(* IEC 61131-3 sources: plcassist-cli/packages/volt-lsp-iec/test-corpus/pro2193/Device/Plc Logic/Application/09 Misc/Library Manager/L_TT1P_TechnologyModules (part 4) *)

(* ---- L_MB1P_TPCALCDIFF.fb ---- *)
FUNCTION_BLOCK L_MB1P_TPCALCDIFF
VAR_INPUT
	XENABLE : BOOL;
	XTPRECEIVED : BOOL;
	LRACTTPPOSIN : LREAL;
	LRSETTPPOSIN : LREAL;
	LRSETMARKDISTANCE : LREAL;
END_VAR
VAR_OUTPUT
	XINITDONE : BOOL;
	XTPRECEIVEDOUT : BOOL;
	LRTPDIFFERENCE : LREAL;
	LRTPDIFFTOTAL : LREAL;
END_VAR
VAR
	XTPRECEIVEDOLD : BOOL;
END_VAR
END_FUNCTION_BLOCK

(* ---- L_MB1P_TPCONVERTTP.fb ---- *)
FUNCTION_BLOCK L_MB1P_TPCONVERTTP
VAR_INPUT
	XENABLE : BOOL;
	XTPRECEIVE : BOOL;
	LRACTTPPOSIN : LREAL;
	LRDELAYACTSET : LREAL;
	LRCYCPOSTPAXIS : LREAL;
	LRCYCPOSTARGETAXIS : LREAL;
	LRCYCLELENGTHTPAXIS : LREAL;
	LRCYCLELENGTHTARGETAXIS : LREAL;
END_VAR
VAR_OUTPUT
	XTPRECEIVED : BOOL;
	LRTPACTPOS : LREAL;
	XERROR : BOOL;
	EERRORID : L_IE1P_Error;
END_VAR
VAR
	LRPOSFIFOX : ARRAY [1..20] OF LREAL := [10(0)];
	LRPOSFIFOREG : ARRAY [1..20] OF LREAL := [10(0)];
	BYCOUNTER : INT := 1;
	LRSTACKDIFFERENCE : LREAL;
	LRTPDELTAINMS : LREAL;
	LRDELTAPCT : LREAL;
	XTPRECEIVEDOLD : BOOL;
	LRPOSDIFFTPAXIS : LREAL;
	IDIRECTION : INT;
	LRACTTPPOSIN_OLD : LREAL;
	XWAIT : BOOL;
	XWAIT_OLD : BOOL;
	LRACTTPPOSIN_INT : LREAL;
	R_TRIG1 : R_TRIG;
	BYCOMPENSATIONCYCLES : BYTE;
	LRDELAYACTSETRESIDUAL : LREAL;
	LRDELTATARGETAXIS : LREAL;
END_VAR
END_FUNCTION_BLOCK

METHOD SEARCHINSTACKNEGATIVE
END_METHOD

METHOD SEARCHINSTACKPOSITIVE
END_METHOD

(* ---- L_MB1P_TPLIMITDIFF.fb ---- *)
FUNCTION_BLOCK L_MB1P_TPLIMITDIFF
VAR_INPUT
	XTPRECEIVED : BOOL;
	LRSETTPDIFFERENCE : LREAL;
	LRSETLIMITMIN : LREAL := -100;
	LRSETLIMITMAX : LREAL := 100;
	LRSETTPWINDOW : LREAL := 2;
END_VAR
VAR_OUTPUT
	XTPRECEIVEDOUT : BOOL;
	XLIMITACTIVE : BOOL;
	XTPINWINDOW : BOOL;
	LRTPDIFFERENCELIM : LREAL;
END_VAR
VAR
	XTPRECEIVEDOLD : BOOL;
	XINITDONE : BOOL;
END_VAR
END_FUNCTION_BLOCK

(* ---- L_MB1P_TPVIRTUALACTPOS.fb ---- *)
FUNCTION_BLOCK L_MB1P_TPVIRTUALACTPOS
VAR_INPUT
	XTPWINDOWOPEN : BOOL;
	XTPRECEIVEDIN : BOOL;
	XMAXTPNOTDETECTED : BOOL;
	LRSETTPPOSIN : LREAL;
	LRACTTPPOSIN : LREAL;
END_VAR
VAR_OUTPUT
	XTPRECEIVEDOUT : BOOL;
	LRACTTPPOS : LREAL;
END_VAR
VAR
	XTPRECEIVEDINOLD : BOOL;
	XFLAGWINDOWOPENANDNOTP : BOOL := FALSE;
	XWINDOWOPENOLD : BOOL;
	XVIRTUALTPACTIVE : BOOL;
END_VAR
END_FUNCTION_BLOCK

(* ---- L_MB1P_WINDERIDENTDIAMETER.fb ---- *)
FUNCTION_BLOCK L_MB1P_WINDERIDENTDIAMETER
VAR_INPUT
	XEXECUTE : BOOL;
	XABORT : BOOL;
	XDANCERMINPOS : BOOL;
	LRACTREELSPEEDIN : LREAL;
	LRACTDANCERPOSIN : LREAL;
	XLINEVELDIAMCALC : BOOL;
	LRSETLINEVELDIAMCALC : LREAL;
	LRMAXDANCERPOS : LREAL;
	LRDANCERMATERIALLENGTH : LREAL;
	LRMAXDIAM : LREAL;
	LRDIAMCALCDIST : LREAL;
	WIDENTDIAMCALCCYCLES : WORD := 1;
	LRTASKCYCLE : LREAL := 0.001;
	LRIDENTVEL : LREAL;
	LRIDENTACC : LREAL;
	LRIDENTDEC : LREAL;
	LRIDENTJERK : LREAL;
END_VAR
VAR_OUTPUT
	XERROR : BOOL;
	EERRORID : WORD;
	XBUSY : BOOL;
	XDONE : BOOL;
	XCOMMANDABORTED : BOOL;
	LRSETREELSPEEDOUT : LREAL;
	LRIDETDIAM : LREAL;
END_VAR
VAR
	WSTATE : WORD;
	LRTASKCYCLE_INT : LREAL := 0.001;
	LRMAXDIAM_INT : LREAL;
	LRREELSPEEDFAKTOR_INT : LREAL;
	LRMAXDANCERPOS_INT : LREAL;
	LRDANCERMATERIALLENGTH_INT : LREAL;
	XLINEVELDIAMCALC_INT : BOOL;
	LRREELSPEEDOUT_INT : LREAL;
	LRACTREELDIST_INT : LREAL;
	LRACTDIST_INT : LREAL;
	LRPROFGENDIST_INT : LREAL;
	LRSETDIST_INT : LREAL;
	LRSETDISTCALCDIAM_INT : LREAL;
	LRPROFGENSTARTPOSIDENTDIAM_INT : LREAL;
	LRPROFGENENDPOSIDENTDIAM_INT : LREAL;
	LRRAMPGENDECDIST : LREAL;
	XRAMPGENHALT : BOOL;
	XIDENTSTARTVALUESVALID : BOOL;
	XIDENTENDVALUESVALID : BOOL;
	LRDANCERPOSSTARTIDENT : LREAL;
	LRDANCERPOSENDIDENT : LREAL;
	LRLINEVELSTARTIDENT : LREAL;
	LRLINEVELENDIDENT : LREAL;
	LRLINEDIST : LREAL;
	LRWNDPOSSTARTIDENT : LREAL;
	LRWNDPOSENDIDENT : LREAL;
	LRIDETNWINDDIST : LREAL;
	XERROR_INVALIDMAXDIAM : BOOL;
	XERROR_INVALIDDANCERMATERIALLENGTH : BOOL;
	XERROR_ACTDANPOSBIGGERMAXDANPOS : BOOL;
	XERROR_ACTDANPOSBIGGERMAXDANPOS_TMP : BOOL;
	XEXECUTE_OLD : BOOL;
	XABORT_OLD : BOOL;
	FB_RAMPGENERATOR1 : L_MC1P_RampGenerator;
END_VAR
END_FUNCTION_BLOCK

METHOD CALL_ERRORHANDLER
END_METHOD

METHOD CALL_FBMETHODS
END_METHOD

METHOD CALL_FB_RAMPGENERATOR
END_METHOD

METHOD CALL_OUTPUT
END_METHOD

METHOD CALL_RESETCOMMANDS
END_METHOD

METHOD CALL_RESETOUTPUT
END_METHOD

METHOD CALL_STATEMACHINE
END_METHOD

(* ---- L_MB1P_WINDERSYNCHRONISELINE.fb ---- *)
FUNCTION_BLOCK L_MB1P_WINDERSYNCHRONISELINE
VAR_INPUT
	XENABLE : BOOL;
	XSYNCLINEVEL : BOOL;
	XLOADSTARTREELSPEED : BOOL;
	LRSTARTREELSPEED : LREAL;
	LRGROUNDREELSPEED : LREAL;
	LRCYCLINEVEL : LREAL := 0;
	LRSETDIAMETER : LREAL;
	LRACC : LREAL := 1000;
	LRDEC : LREAL := 1000;
	LRJERK : LREAL := 100000;
	XMATERIALFEEDING : BOOL := FALSE;
END_VAR
VAR_OUTPUT
	XERROR : BOOL;
	EERRORID : WORD;
	XBUSY : BOOL;
	XSYNCHRONISED : BOOL;
	XACCDECSYNC : BOOL;
	LRSETREELSPEEDOUT : LREAL;
END_VAR
VAR
	WSTATE : WORD;
	LRREELSPEEDOUT_INT : LREAL;
	FB_RAMPGENERATOR1 : L_MC1P_RampGenerator;
	XENABLE_OLD : BOOL;
	XMATERIALFEEDING_OLD : BOOL;
	LRSCALEFAKTOR : LREAL;
	LRSCALEFAKTORABS : LREAL;
	WPARMODE : WORD;
	XTMP : BOOL;
END_VAR
END_FUNCTION_BLOCK

METHOD CALL_ERRORHANDLER
END_METHOD

METHOD CALL_FBMETHODS
END_METHOD

METHOD CALL_FB_RAMPGENERATOR
END_METHOD

METHOD CALL_OUTPUT
END_METHOD

METHOD CALL_RESETCOMMANDS
END_METHOD

METHOD CALL_RESETOUTPUT
END_METHOD

METHOD CALL_SETPARMODE
END_METHOD

METHOD CALL_STATEMACHINE
END_METHOD

(* ---- L_T01S_PHASECORRECTIONVEL.fb ---- *)
FUNCTION_BLOCK L_T01S_PHASECORRECTIONVEL
VAR_INPUT
	XENABLE : BOOL;
	XEXECUTECORRECTION : BOOL;
	LRCYCSETVEL : LREAL;
	LRSETCORRECTION : LREAL;
	LRCORRECTIONDISTANCE : LREAL;
END_VAR
VAR_OUTPUT
	XBUSY : BOOL;
	XCORRECTIONBUSY : BOOL;
	LRSETVELOUT : LREAL;
	LRSETCORRVELOUT : LREAL;
	LRSETPOSCORROUT : LREAL;
	XERROR : BOOL;
	EERRORID : L_IE1P_Error;
END_VAR
VAR
	LRDELTAPOSTOTAL : LREAL;
	LRMASTERDISTANCE : LREAL;
	LRPOSITIONSET : LREAL;
	LRPOSITIONNORMED : LREAL;
	LRPOSITIONOUTNORMED : LREAL;
	LRDELTAPOSCORRECTION : LREAL;
	LRPOSITIONSETOLD : LREAL;
	BYSTEPPER : BYTE;
	LRCORRECTIONDISTANCELOCAL : LREAL;
	LRCORRECTIONLOCAL : LREAL;
	LRDELTAPOSOUT : LREAL;
	XEXECUTECORRECTIONINTERN : BOOL;
	LRTASKCYCLE : LREAL;
	XINIT : BOOL := TRUE;
	INTEGRATE1 : L_USPP_Integrate;
END_VAR
END_FUNCTION_BLOCK

(* ---- L_TF1P_ADDPROFILEPICKANDPLACE.fb ---- *)
FUNCTION_BLOCK L_TF1P_ADDPROFILEPICKANDPLACE
VAR_INPUT
	XENABLE : BOOL;
	XEXECUTEPICKANDPLACE : BOOL;
	XADDPROFILE : BOOL;
	XRESETTARGETSTACK : BOOL;
	XACKPATHHALT : BOOL;
	XABORT : BOOL;
	XNOTCOORDINATEDSTOPALL : BOOL;
	XSINGLESTEP : BOOL;
	LRGRIPPERTIME : LREAL;
	LRPATHJERK : LREAL;
	LRNUMTASKCYCLESBEFOREEXECUTENEXTPROFILE : LREAL := 50;
	XCALCPROFILEMOVEPATH : BOOL;
END_VAR
VAR_OUTPUT
	XERROR : BOOL;
	XWARNING : BOOL;
	EERRORID : L_IE1P_Error;
	XBUSY : BOOL;
	XACTIVE : BOOL;
	XDONE : BOOL;
	XCOMMANDABORTED : BOOL;
	XENDOFPROFILE : BOOL;
	XTARGETSTACKISFULL : BOOL;
	XPATHHOLD : BOOL;
	XPROFILEINPREPARATION : BOOL;
	ISETPROFILENOOUT : INT;
	IPROFILEPOINTPASSED : INT;
	ITARGETPROFILEPOINT : INT;
	ALRTARGETPOSITION : ARRAY [1..12] OF LREAL;
	ESETSEGMENTTYPEOUT : L_MC4P_SegmentType;
	BYNUMOFPOINTSINPROFILE : BYTE;
	BYNUMOFHALTINPROFILE : BYTE;
	LRPATHPREPARATIONTIME : LREAL;
	LRPRECALCPROFILETIME : LREAL;
	XPROFILERESTTIMEVALID : BOOL;
	LRPROFILERESTTIME : LREAL;
	LRINTERRUPTPATHACC : LREAL;
	XLASTACTIVESEGMENT : BOOL;
	XNOACTIVESEGMENT : BOOL;
	XGRIPPERCTRLACTIVE : BOOL;
	XPULSEGRIPPER : BOOL;
	XPATHINTERRUPTOUT : BOOL;
	PAFB_MOVELINABS : POINTER TO ARRAY [1..10] OF L_MC4P_MoveLinearAbsolute_Internal;
	IMOVEPPNO : INT;
	IMOVELINNO : INT;
	PAFB_MOVELINABS1 : POINTER TO ARRAY [1..10] OF L_MC4P_MoveLinearAbsolute_Internal;
	PAFB_MOVELINABS2 : POINTER TO ARRAY [1..10] OF L_MC4P_MoveLinearAbsolute_Internal;
	PAFB_MOVELINABS3 : POINTER TO ARRAY [1..10] OF L_MC4P_MoveLinearAbsolute_Internal;
	XWAITDISABLEMOVECONTPATH : BOOL;
END_VAR
VAR_IN_OUT
	FB_EXTERNALMEMORY : L_MC4P_PickAndPlaceMemory;
	AXESGROUP : AXES_GROUP_KIN;
	ASCPROFILEPAR : ARRAY [1..10] OF L_TT1P_scProfilePar;
END_VAR
VAR
	LWTCHECKSUM_INT : LWORD;
	WSTATE : WORD;
	XSTATEMASHINEBUSY : BOOL;
	XSTATEMASHINEWAIT : BOOL;
	XSTATEMASHINEPATHHOLD : BOOL;
	XMOVEPAPSTATUSSEPPERENTRY : BOOL;
	WMOVEPAPSTATUSSEPPER_OLD : WORD;
	WMOVEPAPSTATUSSEPPER : WORD;
	REQUESTSINFO : DWORD;
	REQUESTSINFO_OLD : DWORD;
	DWRTRIG : DWORD;
	DWFTRIG : DWORD;
	EBUFFERMODEBLENDING_INT : MC_BUFFER_MODE := MC_BUFFER_MODE.mcBlendingLow;
	LRTEMP1 : LREAL;
	LRTEMP2 : LREAL;
	IDX1 : INT;
	IDX2 : INT;
	IDX3 : INT;
	UIDX1 : UINT;
	WDX1 : WORD;
	TTMP1 : TIME;
	WTMP1 : WORD;
	IFOR : INT;
	IFOREND : INT;
	ALRTARGETPOSTMP : ARRAY [1..12] OF LREAL;
	XCOUNTUPPROFILENOOUT : BOOL;
	XERRORINVALIDPROFILE : BOOL;
	XERROR_INVALIDCOORDSYSTEM : BOOL;
	XERROR_INVALIDTARGET : BOOL;
	XERROR_INVALIDPATHPAR : BOOL;
	XWARNING_TARGETSTATCKISFULL : BOOL;
	XWARNING_NOTREADYFORADDPROFILE : BOOL;
	XERROR_FB_MOVEPICKANDPLACE : BOOL;
	EERRORID_FB_MOVEPICKANDPLACE : L_IE1P_Error;
	XERROR_INTERNAL : BOOL;
	XERRORINTERNAL_INVALIDPPFBACTIVE : BOOL;
	WINTERNALERRORID_INT : WORD;
	XSINGLESTEP_LOCK : BOOL;
	LRGRIPPERTIME_LOCK : LREAL;
	XCALLFM : BOOL;
	LRTASKCYCLE : LREAL;
	LRTASKCYCLE_INV : LREAL;
	LRTIMEBEFOREEXECUTENEXTPROFILE : LREAL;
	FB_STACKTARGET : L_MC1P_StackControlArray := STRUCT(iMaxLegth := ciNumOfTargetInArray);
	ALRTARGETGRIPPERTIME : ARRAY [1..ciNumOfTargetInArray] OF LREAL;
	ALRPATHJERK : ARRAY [1..ciNumOfTargetInArray] OF LREAL;
	AXTARGETGRIPPERTIMEVALID : ARRAY [1..ciNumOfTargetInArray] OF BOOL;
	AXSINGLESTEP_INT : ARRAY [1..ciNumOfTargetInArray] OF BOOL;
	XNEWTARGET : BOOL;
	XAXESGROUPNOTREADYFORMOTION : BOOL;
	XNEXTPROFILEVALID : BOOL;
	XMOVEPPPATHINTERRUPTOUT : BOOL;
	IGRIPPERMOVEPPNO : INT;
	XPREPARENEXTPROFILE : BOOL;
	XPATHACTIVE_INT : BOOL;
	XPATHBUSY_INT : BOOL;
	XPATHDONE_INT : BOOL;
	XPATHHOLD_INT : BOOL;
	XPATHHOLDONENDHALT_INT : BOOL;
	XPATHINTERRUPTOUT_INT : BOOL;
	XPATHCOMMANDABORTED_INT : BOOL;
	XCOMMANDABORTED_INT : BOOL;
	XCOMMANDABORTE_INT : BOOL;
	XPROFILEINPREPARATION_INT : BOOL;
	LRPRECALCRESTTIMEALLSEGMENTS_INT : LREAL;
	XPRECALCPROFILERESTTIMEALLSEGMENTSVALID_INT : BOOL;
	XPRECALCPROFILERESTTIMEVALID_INT : BOOL;
	LRPRECALCPROFILERESTTIME_INT : LREAL;
	LRIPOTIME : LREAL;
	LRPATHPREPARATIONTIME_INT : LREAL;
	INUMOFACTIVEPATHSEGMENT_INT : INT;
	ICNTRACKPATHHALT_INT : INT;
	XVALIDSTARTPOS : BOOL;
	XSTARTPOINTINHALT_INT : BOOL;
	ALRSTARTPOS_INT : ARRAY [1..12] OF LREAL;
	ESTARTCOORDSYSTEM_INT : L_MC4P_CoordSystem;
	LRSTARTBLENDINGRADIUS_INT : LREAL;
	XSAVEPROFILE_INT : BOOL;
	ISAVEPROFILEEXECUTED_INT : INT;
	ISAVEPROFILESTACKSTARTPOS_INT : INT;
	ISAVEPROFILESTACKLEGTH_INT : INT;
	FB_STACKMOVEPICKANDPALCE : L_MC1P_StackControlArray := STRUCT(iMaxLegth := ciNumOfFBMovePickAndPlace);
	AIPROFILENOSTATIC : ARRAY [1..ciNumOfFBMovePickAndPlace] OF INT;
	FB_MOVEPICKANDPLACE : ARRAY [1..ciNumOfFBMovePickAndPlace] OF L_MB1P_MovePickAndPlaceState;
	CINUMOFTARGETINARRAY : INT := 10;
	CINUMOFTARGETINARRAYSETWARNING : INT := 8;
	CINUMOFFBMOVEPICKANDPLACE : INT := 3;
	EBUFFERMODEBLENDING : MC_BUFFER_MODE;
	LWTCHECKSUM : LWORD;
END_VAR
END_FUNCTION_BLOCK

METHOD CALL_ALLOCPOINTADR
END_METHOD

METHOD CALL_CALCPROFILETIME
END_METHOD

METHOD CALL_DISABLEMOVECONTPATH
VAR_IN_OUT
	AXESGROUP : AXES_GROUP_KIN;
END_VAR
END_METHOD

METHOD CALL_ERRORHANDLER
END_METHOD

METHOD CALL_FBMETHODS
END_METHOD

METHOD CALL_FB_MOVEPICKANDPLACE
END_METHOD

METHOD CALL_FB_MOVEPICKANDPLACE_STATUS
END_METHOD

METHOD CALL_GRIPPERCONTROL
END_METHOD

METHOD CALL_OUTPUT
END_METHOD

METHOD CALL_REQUESTS_EXT
END_METHOD

METHOD CALL_RESETCOMMANDS
END_METHOD

METHOD CALL_RESETOUTPUT
END_METHOD

METHOD CALL_STATEMACHINE
END_METHOD

METHOD CALL_ABORTPROFILE
END_METHOD

METHOD CALL_READSTARTPOSITION
END_METHOD

METHOD CALL_SAVEPROFILE
END_METHOD

METHOD CALL_TARGETSTAICPOSSTACK
END_METHOD

METHOD CALL_SETPROFILE
END_METHOD

METHOD GET_ALRINTERMEDIANTEPOINT
VAR_IN_OUT
	ALRINTERMEDIANTEPOINT : ARRAY [1..12] OF LREAL;
END_VAR
END_METHOD

METHOD CALL_INIT
END_METHOD

METHOD CALL_S000_CYCLIC
END_METHOD

(* ---- L_TF1P_REGISTERCONTROLBASE.fb ---- *)
FUNCTION_BLOCK L_TF1P_REGISTERCONTROLBASE
VAR_INPUT
	XENABLE : BOOL;
	XSYNCPOS : BOOL;
	LRVELIN : LREAL;
	LRACTSETPOSSLAVE : LREAL;
	XMARKRECEIVE : BOOL;
	ETPMODE : L_TF1P_TpMode;
	LRCYCPOSEXTENCODER : LREAL;
	LRCYCLELENGTHEXTENCODER : LREAL;
	LRACTMARKPOSIN : LREAL;
	XLOADREGPOS : BOOL;
	LRLOADREGPOS : LREAL;
	LRMARKSENSORPOS : LREAL;
	LRMARKDIST : LREAL;
	LRMAXCORRNEG : LREAL;
	LRMAXCORRPOS : LREAL;
	ESOURCEFORCORRWINDOW : L_TT1P_SourceForCorrWindow;
	LRUPPERCORRPOS : LREAL;
	LRLOWERCORRPOS : LREAL;
	DNNUMAXISY : DWORD;
	DNDENAXISY : DWORD;
	XSYNCHRONISED : BOOL;
	LRTPAXISCOMPFACTOR : LREAL;
	LRTPAXISDELAYCYCLE : LREAL;
END_VAR
VAR_OUTPUT
	LRPOSOUT : LREAL;
	LRACTVEL : LREAL;
	XERROR : BOOL;
	WERRORID : WORD;
	XLIMITACTIVE : BOOL;
	LRACTMARKERROR : LREAL;
	LRACTMARKDIST : LREAL;
	XINITDONE : BOOL;
	XCORRACTIVE : BOOL;
	XMARKRECEIVED : BOOL;
	LRREGMARKPOS : LREAL;
	XCORRNEXTCYCLE : BOOL;
END_VAR
VAR_IN_OUT
	MASTERAXIS : AXIS_REF;
	SLAVEAXIS : AXIS_REF;
END_VAR
VAR
	SPEEDTOPOSINTEGRATE : L_MC1P_IntegrateAxis;
	TPLIMITDIFF : L_MB1P_TpLimitDiff;
	FB_ADDOFFSET : L_MC1P_AddOffsetCyclic;
	TPCALCDIFF : L_MC1P_TpCalcDiff;
	CONVERTTPPOSITION : L_TT1P_CalculateTPOnMaterialPos := STRUCT(xNoMarkStack := TRUE);
	DISTCORRECTIONWINDOW : L_MB1P_DistCorrectionWindow;
	LRGEARINGFAKTOR : LREAL := 1.0;
	XERROR_TM : BOOL;
	EERRORID_TM : L_IE1P_Error;
	LRTPDIFFERENCE_INT : LREAL;
	XLOADMARKSENSORPOS_OLD : BOOL;
	XTPRECEIVED_OLD : BOOL;
	LRMARKWINDOWSIZE_INT : LREAL;
	XTPINWINDOW : BOOL;
	LRPOS_INT : LREAL;
	XTPRECEIVEDOUT_INT : BOOL;
	LRTPACTPOSITION_INT : LREAL;
	LRTPDIFFERENCELIM_INT : LREAL;
	LROFFSETPOSCTRL_INT : LREAL;
	LRPOSOUT_INT : LREAL;
	LRVELOUT_INT : LREAL;
	XCORRACTIVE_INT : BOOL;
	XINIT : BOOL := TRUE;
	XTPCORRECTIONACTIVE : BOOL := FALSE;
	LRTPAXISSETPOS : LREAL;
	LRMARKDIST_INT : LREAL;
	XZERO : BOOL;
	XHOMINGDONE : BOOL;
	XSTARTREFERENCEACTIVE : BOOL;
	XHOMINGACTIVE : BOOL := FALSE;
	XMARKDISTCHANGED : BOOL;
	XENABLE_OLD : BOOL;
	XTPRECEIVEDOUT_INTOLD : BOOL;
	XSTARTFIRSTCORRECTION : BOOL;
	LRTPDIFFERENCELIM2_INT : LREAL;
	XCORRECTIONBUSYOLD : BOOL;
	LRTPACTPOSIN_OLD : LREAL;
	LRTPSETPOSIN_OLD : LREAL;
	LRCYCLELENGTH : LREAL;
	ICOUNTER : INT := 0;
	LRSETPOSITIONOLD : LREAL;
	LRCYCLELENGTHTP : LREAL;
	LRTPACTPOSITIONOLD : LREAL;
	L_MB1P_CHECKMODULOOVERRUNSETPOS : L_MB1P_CheckModuloOverrun;
	L_MB1P_CHECKMODULOOVERRUNACTPOS : L_MB1P_CheckModuloOverrun;
	BYCYCLECOUNT_INT : BYTE;
	BYCYCLECOUNTREG_INT : BYTE;
	BYSTATE : BYTE;
	ABYCYCLECOUNT : ARRAY [0..5] OF BYTE;
	BYCYCLECOUNTSUM : BYTE;
	XFIRSTTOUCHPROBE : BOOL := TRUE;
	XCORRBASEDONMASTERPOS_INT : BOOL := FALSE;
	XTPCALCDIFFTPRECEIVEDOLD : BOOL;
	LRTPDIFFERENCECOMP_INT : LREAL;
	LRTPAXISACTPOS : LREAL;
	LRTPAXISACTVELOCITY : LREAL;
	LRTPAXISCYCLELENGTH : LREAL;
	LRCYCREGISTERPOSINT : LREAL;
	LRTPACTPOSITION_ORIGINAL : LREAL;
	LRREGISTERTOUCHPROBEDIFFERENCE : LREAL;
	LRAXISTOUCHPROBEDIFFERENCE : LREAL;
END_VAR
END_FUNCTION_BLOCK

METHOD CALL_CALCACTMARKDIST
END_METHOD

METHOD CALL_CORRECTIONPOS
END_METHOD

METHOD CALL_ENABLEREGISTERCONTROL
END_METHOD

METHOD CALL_ERRORHANDLER
END_METHOD

METHOD CALL_FB
END_METHOD

METHOD CALL_GEARING
END_METHOD

METHOD CALL_INPUT
END_METHOD

METHOD CALL_LIMIT
END_METHOD

METHOD CALL_MARKDISTCHANGE
END_METHOD

METHOD CALL_NOTENABLE
END_METHOD

METHOD CALL_OUTPUT
END_METHOD

METHOD CALL_RESET
END_METHOD

METHOD CALL_TOUCHPROBE
END_METHOD

METHOD CALL_TOUCHPROBESOURCE
END_METHOD

METHOD GET_ACTUALMARKDIST : LREAL
END_METHOD

METHOD GET_CORRREGPOS : LREAL
END_METHOD

METHOD GET_INTEGRATORREGPOS : LREAL
END_METHOD

METHOD GET_MARKERRORUNLIMITED : LREAL
END_METHOD

METHOD GET_MARKPOSITIONINREGISTER : LREAL
END_METHOD

METHOD GET_MARKRECEIVEUNLIMITED : BOOL
END_METHOD

METHOD GET_REGISTERINPUTVEL : LREAL
END_METHOD

METHOD GET_SETVELOCITYREGISTER : LREAL
END_METHOD

METHOD SET_CORRECTIONONMASTERPOS
VAR_INPUT
	XCORRBASEDONMASTER : BOOL;
END_VAR
END_METHOD

(* ---- L_TF1P_REGISTERCONTROLSTATE.fb ---- *)
FUNCTION_BLOCK L_TF1P_REGISTERCONTROLSTATE EXTENDS L_TF1P_RegisterControlBase
VAR_INPUT
	LRACTOFFSETMASTERIN : LREAL;
	LRACTOFFSETSLAVEIN : LREAL;
	XTEACHMARKWINDOW : BOOL;
	LRMARKWINDOWSIZE : LREAL;
	LRSETOFFSETMARKWINDOW : LREAL;
	DWMAXNUMBERVIRTUALMARKS : DWORD;
	LRGEARFACTORCORRGAIN : LREAL;
	LRMAXGEARFACTORCORR : LREAL;
	LRSENSORTOOLDISTANCE : LREAL;
	XGEARFACTORCORR : BOOL;
	XGEARFACTORCORRHOLD : BOOL;
	XENABLETOOLCORRECTION : BOOL;
END_VAR
VAR_OUTPUT
	XMARKWINDOWOPEN : BOOL;
	XMARKOUTOFWINDOW : BOOL;
	XMARKNOTDETECTED : BOOL;
	XMARKWINDOWTEACHED : BOOL;
	LRAVERAGEGEARFACTORCORR : LREAL;
	XGEARFACTORCORRLIMITED : BOOL;
END_VAR
VAR
	MARKWINDOW : L_MB1P_MarkWindowRelative;
	MARKSTACK : L_MB1P_MarkStack;
	TPVIRTUALACTPOS : L_MB1P_TpVirtualActPos;
	LRMARKSTACKLENGTH : LREAL;
	LRTPDIFFERENCELIMITOUT_INT : LREAL;
	XTPRECEIVESTACKOUT_INT : BOOL;
	XTPNOTDETECTED_INT : BOOL;
	XMAXTPNOTDETECTED : BOOL;
	LRGEARFACTORINTEGRATOR : LREAL;
	LRGEARFACTORGAIN : LREAL := 1;
	LRGEARFACTORNUMERATORCORR : LREAL;
	LRGEARFACTORNUMERATORCORRLIMITED : LREAL;
	LRGEARFACTORDENOMINATOR : LREAL;
	LRGEARFACTORNUMERATOR : LREAL;
	LCORRECTIONVELIN : LREAL;
	LRDELTAGEARFACTORCORR : LREAL;
	XTPSENSORTEACHEDOLD : BOOL;
	XTPSENSORTEACHEDATLASTMARK : BOOL;
	XCALCMARKDISTINITIALISED : BOOL;
	XTEACHTPSENSOROLD : BOOL;
	LRTPDEADTIMEDIFF : LREAL;
	XTPRECEIVEDOUTOLD_INT : BOOL;
	XMARKSTACKTPRECEIVEDOUTOLD : BOOL;
	LRTPACTPOSITIONREGISTER_INT : LREAL;
	XTPRECEIVEDOUTREGISTER_INT : BOOL;
	XTPRECEIVEDOUTCALCERROR_INT : BOOL;
	LRTPACTPOSMARKWINDOWIN_INT : LREAL;
	LRMASTERACTPOSITIONOLD_INT : LREAL;
END_VAR
END_FUNCTION_BLOCK

METHOD CALL_AVERAGETPDIFF
END_METHOD

METHOD CALL_CALCACTMARKDIST
END_METHOD

METHOD CALL_CORRECTIONPOS
END_METHOD

METHOD CALL_ENABLEREGISTERCONTROL
END_METHOD

METHOD CALL_ERRORHANDLER
END_METHOD

METHOD CALL_FB
END_METHOD

METHOD CALL_INPUT
END_METHOD

METHOD CALL_LIMIT
END_METHOD

METHOD CALL_MARKDISTCHANGE
END_METHOD

METHOD CALL_MARKREGISTER
END_METHOD

METHOD CALL_MARKWINDOW
END_METHOD

METHOD CALL_NOTENABLE
END_METHOD

METHOD CALL_OUTPUT
END_METHOD

METHOD CALL_RESET
END_METHOD

METHOD CALL_TOUCHPROBE
END_METHOD

METHOD CALL_TOUCHPROBESOURCE
END_METHOD

METHOD CALL_VIRTUALACTPOS
END_METHOD

METHOD GET_ACTMARKERRORLIMITED : LREAL
END_METHOD

METHOD GET_MARKRECEIVEDLIMITED : BOOL
END_METHOD

METHOD GET_MARKWINDOWCOMP : BOOL
END_METHOD

METHOD GET_LRMARKSTACKLENGTH : LREAL
END_METHOD

(* ---- L_TF1P_SYNCDRIVEPOSBASE.fb ---- *)
FUNCTION_BLOCK L_TF1P_SYNCDRIVEPOSBASE
VAR_INPUT
	XENABLE : BOOL;
	LRCYCMASTERPOS : LREAL;
	LRCYCMASTERVEL : LREAL;
	LRCYCMASTERACC : LREAL;
	XLOADSTARTSLAVEPOS : BOOL := FALSE;
	LRSTARTSLAVEPOS : LREAL;
	XLOADGEARBOXPOS : BOOL;
	LRLOADGEARBOXPOS : LREAL;
	DWNUMERATOR : DWORD := 1;
	DWDENOMINATOR : DWORD := 1;
	LRSETOFFSET : LREAL;
END_VAR
VAR_OUTPUT
	XERROR : BOOL;
	EERRORID : L_IE1P_Error;
	XBUSY : BOOL;
	LRSETSLAVEPOSOUT : LREAL;
	LRSETSLAVEVELOUT : LREAL;
	LRSETSLAVEACCOUT : LREAL;
	LRSETGEARBOXPOSOUT : LREAL;
	LROFFSET : LREAL;
END_VAR
VAR_IN_OUT
	MASTERAXIS : AXIS_REF;
	SLAVEAXIS : AXIS_REF;
END_VAR
VAR
	LRSCALING_INT : LREAL := 1;
	LRGEARBOXSTARTPOSOUT_INT : LREAL;
	LRSETMASTERVEL_INT : LREAL;
	LRSETMASTERVEL_OLD : LREAL;
	LRSETMASTERACC_INT : LREAL;
	DWDENOMINATOR_INT : DWORD := 1;
	XENABLE_OLD : BOOL;
	WAXESMODE : WORD;
	ESTATE : L_TF1P_States := L_TF1P_States.INIT;
	ESTATE_OLD : L_TF1P_States := L_TF1P_States.INIT;
	XSTATEENTRY : BOOL;
	XENABLEGEARBOX : BOOL;
	FB_ADDOFFSETCYCLIC : L_MC1P_AddOffsetCyclic;
	FB_GEARBOXPOSITION : L_MB1P_GearboxPosition;
	FB_AXISCONVERTER : L_MC2P.L_MC2P_AxisConverterBase;
	LRLOADGEARBOXPOS_INT : LREAL;
	LRSETGEARBOXPOSOUT_INT : LREAL;
	LRSETGEARBOXPOSOUT_OLD : LREAL;
END_VAR
END_FUNCTION_BLOCK

METHOD CALL_AXESMODE
END_METHOD

METHOD CALL_ERRORHANDLER
END_METHOD

METHOD CALL_FBMETHODS
END_METHOD

METHOD CALL_FBMETHODS_FMDISABLE
END_METHOD

METHOD CALL_FB_ADDOFFSETCYCLIC
END_METHOD

METHOD CALL_FB_ADDOFFSETCYCLIC_INPUT
END_METHOD

METHOD CALL_FB_AXISCONVERTER
END_METHOD

METHOD CALL_FB_AXISCONVERTER_INPUT
END_METHOD

METHOD CALL_FB_GEARBOXPOSITION
END_METHOD

METHOD CALL_FB_GEARBOXPOSITION_INPUT
END_METHOD

METHOD CALL_FB_GEARBOXPOSITION_LOADGEARBOXPOS
END_METHOD

METHOD CALL_LOADSLAVESTARTPOS
END_METHOD

METHOD CALL_OUTPUT
END_METHOD

METHOD CALL_OUTPUT_OFFSET
END_METHOD

METHOD CALL_OUTPUT_SETSLAVEOUT
END_METHOD

METHOD CALL_RESETCOMMANDS
END_METHOD

METHOD CALL_RESETFM
END_METHOD

METHOD CALL_RESETOUTPUT
END_METHOD

METHOD CALL_STATEMASHINE
END_METHOD

METHOD CALL_S000_CYCLIC
END_METHOD

METHOD CALL_S001_INIT
END_METHOD

METHOD CALL_S010_READY
END_METHOD

METHOD CALL_S200_SYNCHRON
END_METHOD

METHOD CALL_S998_ERROR
END_METHOD

(* ---- L_TF1P_SYNCDRIVEPOSHIGH.fb ---- *)
FUNCTION_BLOCK L_TF1P_SYNCDRIVEPOSHIGH EXTENDS L_TF1P_SyncDrivePosState
VAR_INPUT
	XSYNCINSTANT : BOOL;
	XSYNCPOSRESTORE : BOOL;
	XLOADOFFSET : BOOL;
	EOFFSETDIRECTION : L_TF1P_Direction;
	EOFFSETPROFILETYPE : L_TF1P_ProfileType := 0;
	LROFFSETVELPOS : LREAL := 100.0;
	LROFFSETVELNEG : LREAL := 100.0;
	LROFFSETACCDEC : LREAL := 1000.0;
	ESYNCDIRECTION : L_TF1P_SyncDirection := L_TF1P_SyncDirection.mcShortestWay;
	ESYNCMODE : L_TF1P_SyncMode := L_TF1P_SyncMode.ramp_dist;
	LRSYNCINTIME : LREAL := 5;
	LRSYNCOUTTIME : LREAL := 5;
	LRSYNCVEL : LREAL := 100;
	LRSYNCACC : LREAL := 1000.0;
	LRSYNCDEC : LREAL := 1000.0;
	LRSYNCJERK : LREAL := 10000000000.0;
	XLOADCLUTCHOFFSET : BOOL := FALSE;
	LRLOADCLUTCHOFFSET : LREAL := 0;
END_VAR
VAR_OUTPUT
	XSETOFFSETBUSY : BOOL;
	XSETOFFSETDONE : BOOL;
	LROFFSETSYNCPOS : LREAL;
END_VAR
VAR
	LRLOADOFFSET_INT : LREAL := 0;
	XSYNCINSTANT_OLD : BOOL;
	FB_SIMPLEPOSSETOFFSETSLAVE : L_MB1P_SimplePosSetOffset;
	FB_SIMPLEPOSSETOFFSETSYNC : L_MB1P_SimplePosSetOffset;
	LRSYNCOFFSET : LREAL;
END_VAR
END_FUNCTION_BLOCK

METHOD CALL_ERRORHANDLER
END_METHOD

METHOD CALL_FBMETHODS
END_METHOD

METHOD CALL_FBMETHODS_FMDISABLE
END_METHOD

METHOD CALL_FB_ADDOFFSETCYCLIC_INPUT
END_METHOD

METHOD CALL_FB_CLUTCHEXTENDEDBASE_INPUT
END_METHOD

METHOD CALL_FB_SIMPLEPOSSETOFFSETSLAVE
END_METHOD

METHOD CALL_FB_SIMPLEPOSSETOFFSETSLAVE_INPUT
END_METHOD

METHOD CALL_FB_SIMPLEPOSSETOFFSETSYNC
END_METHOD

METHOD CALL_FB_SIMPLEPOSSETOFFSETSYNC_INPUT
END_METHOD

METHOD CALL_OUTPUT
END_METHOD

METHOD CALL_OUTPUT_OFFSET
END_METHOD

METHOD CALL_OUTPUT_SIMPLEPOS
END_METHOD

METHOD CALL_RESETCOMMANDS
END_METHOD

METHOD CALL_RESETOUTPUT
END_METHOD

METHOD CALL_SIMPLEPOS_OFFSET
END_METHOD

METHOD CALL_S001_INIT
END_METHOD

(* ---- L_TF1P_SYNCDRIVEPOSSTATE.fb ---- *)
FUNCTION_BLOCK L_TF1P_SYNCDRIVEPOSSTATE EXTENDS L_TF1P_SyncDrivePosBase
VAR_INPUT
	XSYNCPOS : BOOL;
	XSYNCOUTINSTANT : BOOL;
	XTRIMPOS : BOOL;
	XTRIMNEG : BOOL;
	XRESETTRIM : BOOL;
	LRCYCSLAVEPOS : LREAL;
	LRCYCSLAVEVEL : LREAL;
	LRCYCSLAVEACC : LREAL;
	LRTRIMVELPOS : LREAL := 10.0;
	LRTRIMVELNEG : LREAL := 10.0;
	LRTRIMACC : LREAL := 100.0;
	LRTRIMDEC : LREAL := 100.0;
	XLOADTRIMOFFSET : BOOL;
	LRLOADTRIMOFFSET : LREAL := 0;
	LRSLAVESYNCOUTPOS : LREAL;
	LRSLAVESYNCINDIST : LREAL := 90;
	LRSLAVESYNCOUTDIST : LREAL := 90;
	LRSYNCOUTINSTANTDEC : LREAL := 10000;
END_VAR
VAR_OUTPUT
	XSYNCOUTDONE : BOOL;
	XSYNCHRONISED : BOOL;
	XACCDECSYNC : BOOL;
	XTRIMBUSY : BOOL;
	LRSETTRIMVELOUT : LREAL;
	LROFFSETTRIM : LREAL;
	LROFFSETTOTAL : LREAL;
	LRSETCLUTCHPOS : LREAL;
	LRSETCLUTCHVEL : LREAL;
	LRSETCLUTCHACC : LREAL;
END_VAR
VAR
	LRLOADTRIMOFFSET_INT : LREAL := 0;
	LRSYNCOUTINSTANTDEC_INT : LREAL := 100000;
	LRSETINTEGRATETRIMVELPOSOUT_INT : LREAL;
	XSYNCPOS_OLD : BOOL;
	XRESETTRIM_OLD : BOOL;
	FB_LDMPOTTRIMVEL : L_MC1P_MPot;
	FB_INTEGRATETRIMVEL : L_MC1P_IntegrateAxis;
	FB_CLUTCHEXTENDEDBASE : L_MB1P_ClutchExtendedBase;
END_VAR
END_FUNCTION_BLOCK

METHOD CALL_ERRORHANDLER
END_METHOD

METHOD CALL_FBMETHODS
END_METHOD

METHOD CALL_FBMETHODS_FMDISABLE
END_METHOD

METHOD CALL_FBMETHODS_TRIMVEL
END_METHOD

METHOD CALL_FB_ADDOFFSETCYCLIC_INPUT
END_METHOD

METHOD CALL_FB_CLUTCHEXTENDEDBASE
END_METHOD

METHOD CALL_FB_CLUTCHEXTENDEDBASE_INPUT
END_METHOD

METHOD CALL_FB_CLUTCHEXTENDEDBASE_INPUTMASTER
END_METHOD

METHOD CALL_FB_CLUTCHEXTENDEDBASE_INPUTSLAVE
END_METHOD

METHOD CALL_FB_INTEGRATETRIMVEL
END_METHOD

METHOD CALL_FB_INTEGRATETRIMVEL_INPUT
END_METHOD

METHOD CALL_FB_INTEGRATETRIMVEL_LOADVALUE
END_METHOD

METHOD CALL_FB_LDMPOTTRIMVEL
END_METHOD

METHOD CALL_FB_LDMPOTTRIMVEL_INPUT
END_METHOD

METHOD CALL_LOADSLAVESTARTPOS
END_METHOD

METHOD CALL_OUTPUT
END_METHOD

METHOD CALL_OUTPUT_CLUTCHSTATE
END_METHOD

METHOD CALL_OUTPUT_OFFSET
END_METHOD

METHOD CALL_OUTPUT_SETSLAVEOUT
END_METHOD

METHOD CALL_RESETCOMMANDS
END_METHOD

METHOD CALL_RESETOUTPUT
END_METHOD

METHOD CALL_S000_CYCLIC
END_METHOD

METHOD CALL_S001_INIT
END_METHOD

METHOD CALL_S200_SYNCHRON
END_METHOD

(* ---- L_TF1P_SYNCDRIVEREGCTRL.fb ---- *)
FUNCTION_BLOCK L_TF1P_SYNCDRIVEREGCTRL EXTENDS L_TF1P_SyncDrivePosHigh
VAR_INPUT
	XMASTERTRIM : BOOL;
	XMODULOAXISISREQUIRED : BOOL;
	EOFFSETMASTERDIRECTION : L_TF1P_Direction;
	EOFFSETMASTERPROFILETYPE : L_TF1P_ProfileType := 0;
	LROFFSETMASTERMAXVELPOS : LREAL := 100.0;
	LROFFSETMASTERMAXVELNEG : LREAL := 100.0;
	LROFFSETMASTERACCDEC : LREAL := 1000.0;
	ETRIMMODE : L_TF1P_TrimMode := 0;
	LRTRIMDIST : LREAL;
	LRSETOFFSETMASTER : LREAL;
	XLOADOFFSETMASTER : BOOL;
END_VAR
VAR_OUTPUT
	LROFFSETMASTER : LREAL;
	LROFFSETSLAVE : LREAL;
END_VAR
VAR
	LRSETOFFSETMASTER_INT : LREAL;
	LRTRIMDIST_INT : LREAL;
	XTRIMPOS_OLD : BOOL;
	XTRIMNEG_OLD : BOOL;
	XTRIMVEL : BOOL;
	LRTRIMOFFSETDIST : LREAL;
	LRLOADOFFSETMASTER_INT : LREAL := 0;
	FB_SIMPLEPOSSETOFFSETMASTER : L_MB1P_SimplePosSetOffset;
	FB_SIMPLEPOSTRIMDIST : L_MB1P_SimplePosSetOffset;
	FB_ADDOFFSETCYCLICMASTER : L_MC1P_AddOffsetCyclic;
END_VAR
END_FUNCTION_BLOCK

METHOD CALL_ERRORHANDLER
END_METHOD

METHOD CALL_FBMETHODS
END_METHOD

METHOD CALL_FBMETHODS_FMDISABLE
END_METHOD

METHOD CALL_FBMETHODS_TRIMVEL
END_METHOD

METHOD CALL_FBMETHODS_TRIMVEL_MASTER
END_METHOD

METHOD CALL_FBMETHODS_OLD
END_METHOD

METHOD CALL_FB_ADDOFFSETCYCLICMASTER
END_METHOD

METHOD CALL_FB_ADDOFFSETCYCLICMASTER_INPUT
END_METHOD

METHOD CALL_FB_ADDOFFSETCYCLIC_INPUT
END_METHOD

METHOD CALL_FB_AXISCONVERTER_INPUT
END_METHOD

METHOD CALL_FB_GEARBOXPOSITION_INPUT
END_METHOD

METHOD CALL_FB_INTEGRATETRIMVEL_LOADVALUE
END_METHOD

METHOD CALL_FB_LDMPOTTRIMVEL_INPUT
END_METHOD

METHOD CALL_FB_SIMPLEPOSSETOFFSETMASTER
END_METHOD

METHOD CALL_FB_SIMPLEPOSSETOFFSETMASTER_INPUT
END_METHOD

METHOD CALL_FB_SIMPLEPOSTRIMDIST
END_METHOD

METHOD CALL_FB_SIMPLEPOSTRIMDIST_INPUT
END_METHOD

METHOD CALL_LOADSLAVESTARTPOS
END_METHOD

METHOD CALL_OUTPUT
END_METHOD

METHOD CALL_OUTPUT_OFFSET
END_METHOD

METHOD CALL_RESETCOMMANDS
END_METHOD

METHOD CALL_TRIMMODE
END_METHOD

METHOD GET_LRCLUTCHPOSIN : LREAL
END_METHOD

METHOD GET_LROFFSETADDOFFSETCYCLIC : LREAL
END_METHOD

METHOD GET_LRXGEARBOXPOSITION : LREAL
END_METHOD

METHOD GET_LRYGEARBOXPOSITION : LREAL
END_METHOD

METHOD CALL_S001_INIT
END_METHOD

(* ---- L_TF1P_SYNCDRIVEVELBASE.fb ---- *)
FUNCTION_BLOCK L_TF1P_SYNCDRIVEVELBASE
VAR_INPUT
	XENABLE : BOOL;
	LRCYCMASTERVEL : LREAL;
	LRSETOFFSETVEL : LREAL;
	DWMODE : DWORD := 1;
	LRCOUPLINGX : LREAL := 1.0;
	LRCOUPLINGY : LREAL := 1.0;
END_VAR
VAR_OUTPUT
	XERROR : BOOL;
	EERRORID : L_IE1P_Error;
	XBUSY : BOOL;
	LRSETSLAVEVELOUT : LREAL;
	LROFFSET : LREAL;
END_VAR
VAR_IN_OUT
	MASTERAXIS : AXIS_REF;
	SLAVEAXIS : AXIS_REF;
END_VAR
VAR
	XENABLE_OLD : BOOL;
	ESTATE : L_TF1P_States := L_TF1P_States.INIT;
	ESTATE_OLD : L_TF1P_States := L_TF1P_States.INIT;
	XSTATEENTRY : BOOL;
	FB_CONVAXISV : L_MC2P_ConvAxisV;
END_VAR
END_FUNCTION_BLOCK

METHOD CALL_ERRORHANDLER
END_METHOD

METHOD CALL_FBMETHODS
END_METHOD

METHOD CALL_FBMETHODS_FMDISABLE
END_METHOD

METHOD CALL_FB_CONVAXISV
END_METHOD

METHOD CALL_FB_CONVAXISV_INPUT
END_METHOD

METHOD CALL_OUTPUT
END_METHOD

METHOD CALL_OUTPUT_OFFSET
END_METHOD

METHOD CALL_OUTPUT_SETSLAVEOUT
END_METHOD

METHOD CALL_RESETCOMMANDS
END_METHOD

METHOD CALL_RESETFM
END_METHOD

METHOD CALL_RESETOUTPUT
END_METHOD

METHOD CALL_STATEMASHINE
END_METHOD

METHOD GET_MP_LRSETCLUTCHVEL : LREAL
END_METHOD

METHOD GET_CONVAXISV_OUT : LREAL
END_METHOD

METHOD CALL_S000_CYCLIC
END_METHOD

METHOD CALL_S001_INIT
END_METHOD

METHOD CALL_S010_READY
END_METHOD

METHOD CALL_S998_ERROR
END_METHOD

(* ---- L_TF1P_SYNCDRIVEVELHIGH.fb ---- *)
FUNCTION_BLOCK L_TF1P_SYNCDRIVEVELHIGH EXTENDS L_TF1P_SyncDriveVelState
VAR_INPUT
	XLOADOFFSET : BOOL;
	LROFFSETVELACC : LREAL := 10.0;
	LROFFSETVELDEC : LREAL := 10.0;
	LROFFSETVELJERK : LREAL := 1.0;
	XLOADGROUNDVEL : BOOL;
	LRSETGROUNDVEL : LREAL;
	LRGROUNDVELACC : LREAL := 10.0;
	LRGROUNDVELDEC : LREAL := 10.0;
	LRGROUNDVELJERK : LREAL := 1.0;
END_VAR
VAR_OUTPUT
	XSYNCHRONISEDGROUNDVEL : BOOL;
	XACCDECGROUNDVEL : BOOL;
END_VAR
VAR
	LRSETGROUNDVEL_INT : LREAL;
	FB_RAMPGENOFFSET : L_MC1P_RampGenerator;
	FB_RAMPGENGROUNDVEL : L_MC1P_RampGenerator;
END_VAR
END_FUNCTION_BLOCK

METHOD CALL_ERRORHANDLER
END_METHOD

METHOD CALL_FBMETHODS
END_METHOD

METHOD CALL_FB_CLUTCHV_INPUT
END_METHOD

METHOD CALL_FB_RAMPGENGROUNDVEL
END_METHOD

METHOD CALL_FB_RAMPGENGROUNDVEL_INPUT
END_METHOD

METHOD CALL_FB_RAMPGENOFFSET
END_METHOD

METHOD CALL_FB_RAMPGENOFFSET_INPUT
END_METHOD

METHOD CALL_OUTPUT
END_METHOD

METHOD CALL_OUTPUT_OFFSET
END_METHOD

METHOD CALL_RESETCOMMANDS
END_METHOD

METHOD CALL_RESETOUTPUT
END_METHOD

(* ---- L_TF1P_SYNCDRIVEVELSTATE.fb ---- *)
FUNCTION_BLOCK L_TF1P_SYNCDRIVEVELSTATE EXTENDS L_TF1P_SyncDriveVelBase
VAR_INPUT
	XSYNCVEL : BOOL;
	XSYNCOUTVELINSTANT : BOOL;
	XTRIMPOS : BOOL;
	XTRIMNEG : BOOL;
	LRTRIMVELPOS : LREAL := 10.0;
	LRTRIMVELNEG : LREAL := 10.0;
	LRTRIMACC : LREAL := 10.0;
	LRTRIMDEC : LREAL := 10.0;
	XSYNCVELRESET : BOOL;
	LRSYNCINACC : LREAL := 10.0;
	LRSYNCOUTACC : LREAL := 10.0;
	LRSYNCOUTINSTANTDEC : LREAL := 100.0;
	LRSYNCJERK : LREAL := 1.0;
	XAVOIDVELGAPS : BOOL;
END_VAR
VAR_OUTPUT
	LROFFSETTRIM : LREAL;
	LROFFSETTOTAL : LREAL;
	XTRIMBUSY : BOOL;
	XSYNCHRONISED : BOOL;
	XACCDECSYNC : BOOL;
	XSYNCOUTDONE : BOOL;
END_VAR
VAR
	XACCDECSYNC_OLD : BOOL;
	XSYNCVEL_OLD : BOOL;
	XOPEN_OLD : BOOL;
	XINITFB_CLUTCHV : BOOL;
	FB_CLUTCHV : L_MC2P_ClutchVelocity;
	FB_TRIMSPEED : L_MC1P_MPot;
END_VAR
END_FUNCTION_BLOCK

METHOD CALL_ERRORHANDLER
END_METHOD

METHOD CALL_FBMETHODS
END_METHOD

METHOD CALL_FBMETHODS_FMDISABLE
END_METHOD

METHOD CALL_FB_CLUTCHV
END_METHOD

METHOD CALL_FB_CLUTCHV_INPUT
END_METHOD

METHOD CALL_FB_CLUTCHV_PAR
END_METHOD

METHOD CALL_FB_CONVAXISV_INPUT
END_METHOD

METHOD CALL_FB_TRIMSPEED
END_METHOD

METHOD CALL_FB_TRIMSPEED_INPUT
END_METHOD

METHOD CALL_OUTPUT
END_METHOD

METHOD CALL_OUTPUT_OFFSET
END_METHOD

METHOD CALL_OUTPUT_SETSLAVEOUT
END_METHOD

METHOD CALL_RESETCOMMANDS
END_METHOD

METHOD CALL_RESETOUTPUT
END_METHOD

METHOD GET_MP_LRSETCLUTCHVEL : LREAL
END_METHOD

METHOD CALL_S001_INIT
END_METHOD

(* ---- L_TF1P_WINDERJOGGING.fb ---- *)
FUNCTION_BLOCK L_TF1P_WINDERJOGGING
VAR_INPUT
	XJOGLINEPOS : BOOL;
	XJOGLINENEG : BOOL;
	LRSETDIAMETER : LREAL;
	LRJOGLINEACC : LREAL := 10000;
	LRJOGLINEDEC : LREAL := 10000;
	LRJOGLINEVEL : LREAL := 7200;
	XMATERIALFEEDING : BOOL := FALSE;
	XFOLLOWERACTIVE : BOOL;
END_VAR
VAR_OUTPUT
	XERROR : BOOL;
	EERRORID : WORD;
	XBUSY : BOOL;
	XDONE : BOOL;
	XENABLESPEEDFOLLOWER : BOOL;
	LRSETREELSPEED : LREAL;
END_VAR
VAR
	ETMSTATE_INT : L_TF1P_States := L_TF1P_States.INIT;
	LRSETVELOCITY : LREAL;
	L_D94A_SDRAMPGENERATOR1 : L_MC1P_RampGenerator;
END_VAR
END_FUNCTION_BLOCK

METHOD CALL_FB
END_METHOD

METHOD CALL_STATEMACHINE
END_METHOD

METHOD CALL_S001_INIT
END_METHOD

METHOD CALL_S002_READY
END_METHOD

METHOD CALL_S011_JOGPOS
END_METHOD

METHOD CALL_S012_JOGNEG
END_METHOD

METHOD S001_INIT
END_METHOD

METHOD S002_READY
END_METHOD

METHOD S011_JOGPOS
END_METHOD

METHOD S012_JOGNEG
END_METHOD

(* ---- L_TF1P_XYCONTROLLER.fb ---- *)
FUNCTION_BLOCK L_TF1P_XYCONTROLLER
VAR_INPUT
	XEXECUTEX : BOOL;
	XEXECUTEY : BOOL;
	EMODE : L_TT1P_XYMode := L_TT1P_XYMode.NotCoordinated;
	XACITVATEBUFFERRANGE : BOOL;
	SCPROFILEDATAX : L_TT1P_XYProfileData;
	SCPROFILEDATAY : L_TT1P_XYProfileData;
	SCMINLIMITSX : L_TT1P_XYLimits;
	SCMINLIMITSY : L_TT1P_XYLimits;
	SCBUFFERDATA : L_TT1P_XYBufferData;
END_VAR
VAR_OUTPUT
	XBUSY : BOOL;
	XACTIVE : BOOL;
	XDONE : BOOL;
	XERROR : BOOL;
	EERRORID : L_IE1P_Error;
	XACTIVEX : BOOL;
	XACTIVEY : BOOL;
	XDONEX : BOOL;
	XDONEY : BOOL;
	XCOMMANDABORTEDX : BOOL;
	XCOMMANDABORTEDY : BOOL;
END_VAR
VAR_IN_OUT
	AXISX : AXIS_REF;
	AXISY : AXIS_REF;
END_VAR
VAR
	SINSTANCESTR : STRING;
	DWINSTANCEX : POINTER TO BYTE;
	DWINSTANCEY : POINTER TO BYTE;
	FBBASEX : L_MC1P_Template;
	FBBASEY : L_MC1P_Template;
	FBMBX : L_MC1P_MoveBasic;
	FBMBY : L_MC1P_MoveBasic;
	EFUNCTIONTYPX : L_MC1P_TypeFunction;
	EFUNCTIONTYPY : L_MC1P_TypeFunction;
	XERRORX_INT : BOOL;
	EERRORIDX_INT : L_IE1P_Error;
	XERRORY_INT : BOOL;
	EERRORIDY_INT : L_IE1P_Error;
	XBUSYX_INT : BOOL;
	XBUSYY_INT : BOOL;
	XACTIVEX_INT : BOOL;
	XACTIVEY_INT : BOOL;
	XWAITSTARTX : BOOL;
	XWAITSTARTY : BOOL;
	XEXECUTEXOLD : BOOL;
	XEXECUTEYOLD : BOOL;
	XEXECUTEY_INT : BOOL;
	XEXECUTEX_INT : BOOL;
	XENABLECALCULATION : BOOL;
	XWAITPROFILEGENERATIONX : BOOL;
	XWAITPROFILEGENERATIONY : BOOL;
	XSTARTMANIPULATION : BOOL;
	XRESETOUTPUTX : BOOL := TRUE;
	XRESETOUTPUTY : BOOL := TRUE;
	XDONEX_INT : BOOL;
	XDONEY_INT : BOOL;
	EMODE_INT : L_TT1P_XYMode := L_TT1P_XYMode.NotCoordinated;
	SCACTMINLIMITSX : L_TT1P_XYLimits;
	SCACTMINLIMITSY : L_TT1P_XYLimits;
	SCACTPROFILEDATAX : L_TT1P_XYProfileData;
	SCACTPROFILEDATAY : L_TT1P_XYProfileData;
	LRTIMESTART : ARRAY [1..2] OF LREAL;
	XUPDATETIMESTART : ARRAY [1..2] OF BOOL;
	LRTIMECOUNTER : LREAL;
	LRCORRECTTIMEBASEX : LREAL;
	LRCORRECTTIMEBASEY : LREAL;
	SCACTBUFFERDATA : L_MC1P_BufferData;
	XACHSE : WORD := 1;
	YACHSE : WORD := 2;
	C_NOTCOORDINATED : WORD := 0;
	C_SYNCSTARTSTOP : WORD := 1;
	C_ASYNCSTARTSYNCSTOP : WORD := 2;
	C_SYNCSTARTASYNCSTOP : WORD := 3;
	C_ASYNCSTARTSYNCSTOPTIMEOPT : WORD := 4;
	C_SYNCSTARTASYNCSTOPTIMEOPT : WORD := 5;
	ALRPROFILEXACC : ARRAY [0..8] OF LREAL;
	ALRPROFILEXBUFFPOS : ARRAY [0..8] OF LREAL;
	ALRPROFILEXJERK : ARRAY [0..8] OF LREAL;
	ALRPROFILEXPOS : ARRAY [0..8] OF LREAL;
	ALRPROFILEXTIME : ARRAY [0..8] OF LREAL;
	ALRPROFILEXVEL : ARRAY [0..8] OF LREAL;
	ALRPROFILEYACC : ARRAY [0..8] OF LREAL;
	ALRPROFILEYJERK : ARRAY [0..8] OF LREAL;
	ALRPROFILEYPOS : ARRAY [0..8] OF LREAL;
	ALRPROFILEYTIME : ARRAY [0..8] OF LREAL;
	ALRPROFILEYVEL : ARRAY [0..8] OF LREAL;
	XPROFILEDATAXVALID : BOOL;
	XPROFILEDATAYVALID : BOOL;
END_VAR
END_FUNCTION_BLOCK

METHOD CALCULATEMODES
VAR_IN_OUT
	AXISX : AXIS_REF;
	AXISY : AXIS_REF;
END_VAR
END_METHOD

METHOD CHECKINPUTDATAX : BOOL
VAR_IN_OUT
	AXISX : AXIS_REF;
END_VAR
END_METHOD

METHOD CHECKINPUTDATAY : BOOL
VAR_IN_OUT
	AXISY : AXIS_REF;
END_VAR
END_METHOD

METHOD MANIPULATEPROFILEDATA : BOOL
VAR_INPUT
	LRTIMEBASE : LREAL;
	DNCALCMODE : DINT;
END_VAR
VAR_OUTPUT
	XMINVEL : BOOL;
END_VAR
VAR_IN_OUT
	SCPROFILEDATA : L_MC1P_ProfileData;
	SCPROFILEPARAMETER : L_MC1P_ProfileParameter;
	SCMINLIMITS : L_TT1P_XYLimits;
END_VAR
END_METHOD

METHOD MANIPULATEPROFILEDATABUFFER : BOOL
VAR_INPUT
	LRTIMEBASE : LREAL;
	DNCALCMODE : DINT;
	LRBUFFTIMECONST : LREAL;
	LRBUFFTIMEDEC : LREAL;
	LRBUFFTIMEACC : LREAL;
	LRDISTANCE : LREAL;
END_VAR
VAR_OUTPUT
	XMINACC : BOOL;
	XMINDEC : BOOL;
	XMINVEL : BOOL;
END_VAR
VAR_IN_OUT
	SCPROFILEDATA : L_MC1P_ProfileData;
	SCPROFILEPARAMETER : L_MC1P_ProfileParameter;
	SCMINLIMITS : L_TT1P_XYLimits;
END_VAR
END_METHOD

METHOD MANIPULATEPROFILEDATASIMPLE : BOOL
VAR_INPUT
	LRTIMEFACTOR : LREAL;
	LRTIMEBASE : LREAL;
END_VAR
VAR_OUTPUT
	XMINACC : BOOL;
	XMINDEC : BOOL;
	XMINVEL : BOOL;
END_VAR
VAR_IN_OUT
	SCPROFILEDATA : L_MC1P_ProfileData;
	SCPROFILEPARAMETER : L_MC1P_ProfileParameter;
	SCMINLIMITS : L_TT1P_XYLimits;
END_VAR
END_METHOD

METHOD MANIPULATEPROFILEDATASIMPLEVEL : BOOL
VAR_INPUT
	LRTIMEBASE : LREAL;
	LRDELTAPOS : LREAL;
END_VAR
VAR_OUTPUT
	XMINVEL : BOOL;
END_VAR
VAR_IN_OUT
	SCPROFILEPARAMETER : L_MC1P_ProfileParameter;
	SCMINLIMITS : L_TT1P_XYLimits;
END_VAR
END_METHOD

METHOD MANIPULATEPROFILEDATAVEL : BOOL
VAR_INPUT
	LRTIMEBASE : LREAL;
	LRDISTANCE : LREAL;
END_VAR
VAR_OUTPUT
	XMINVEL : BOOL;
END_VAR
VAR_IN_OUT
	SCPROFILEDATA : L_MC1P_ProfileData;
	SCPROFILEPARAMETER : L_MC1P_ProfileParameter;
	SCMINLIMITS : L_TT1P_XYLimits;
END_VAR
END_METHOD

METHOD UPDATELIMITS
VAR_IN_OUT
	SCLIMITS : L_TT1P_XYLimits;
	SCLIMITSORIG : L_TT1P_XYLimits;
	SCPROFILEDATA : L_MC1P_ProfileData;
END_VAR
END_METHOD

METHOD FB_INIT : BOOL
VAR_INPUT
	BINITRETAINS : BOOL;
	BINCOPYCODE : BOOL;
END_VAR
END_METHOD

METHOD CALCSQRT : LREAL
VAR_INPUT
	ARG1 : LREAL;
END_VAR
END_METHOD

METHOD CONVERTMODE : WORD
VAR_INPUT
	EMODE : L_TT1P_XYMode;
	XLIFTUP : BOOL;
END_VAR
END_METHOD

METHOD OVERRIDEHANDLING
VAR_INPUT
	XCALCVEL : BOOL;
	XCALCACC : BOOL;
END_VAR
VAR_IN_OUT
	AXIS : AXIS_REF;
	SCPROFILEPARAMETER : L_MC1P_ProfileParameter;
END_VAR
END_METHOD

(* ---- L_TT1P_BASICMOTIONBASE.fb ---- *)
FUNCTION_BLOCK L_TT1P_BASICMOTIONBASE
VAR_INPUT
	XENABLEINTERNALCONTROL : BOOL;
	XENABLE : BOOL;
	SCCTRLABC : scCtrl_ABC;
	XRESETERROR : BOOL;
	XREGULATORON : BOOL;
	XSTOP : BOOL;
	XHALT : BOOL;
	SCPAR : L_TT1P_scPar_BasicMotionBase;
	XJOGPOS : BOOL;
	XJOGNEG : BOOL;
	XHOMEEXECUTE : BOOL;
	XHOMEABSSWITCH : BOOL;
	XMOVEVELEXECUTE : BOOL;
	XMOVEABSEXECUTE : BOOL;
	XMOVERELEXECUTE : BOOL;
	LRSETPOS_DIST : LREAL;
	XDISABLESWLIMIT : BOOL;
	LROVERRIDE : LREAL := 1.0;
	LROVERRIDEACC : LREAL := 1.0;
	LROVERRIDEJERK : LREAL := 1.0;
END_VAR
VAR_OUTPUT
	XINTERNALCONTROLACTIVE : BOOL;
	ETMSTATE : L_TT1P_States := L_TT1P_States.INIT;
	SCSTATUSABC : scStatus_ABC;
	XERROR : BOOL;
	XWARNING : BOOL;
	EERRORID : L_IE1P_Error;
	SCERRORINFO : L_TT1P_scErrorInfo;
	XAXISENABLED : BOOL;
	XAXISREADY : BOOL;
	XISHOMED : BOOL;
	XDONE : BOOL;
	XBUSY : BOOL;
	XCOMMANDABORTED : BOOL;
	XINPOSITION : BOOL;
	XHWLIMITSWITCHNEG : BOOL;
	XHWLIMITSWITCHPOS : BOOL;
	XSWLIMITENABLED : BOOL;
	XSWLIMITSWITCHNEG : BOOL;
	XSWLIMITSWITCHPOS : BOOL;
	EAXISSTATE : L_MC1P_AXIS_STATE;
	ECONTROLMODE : L_MC1P_ControlMode;
	LRACTVEL : LREAL;
	LRACTPOS : LREAL;
	LRSETPOSOUT : LREAL;
	LRSETVELOUT : LREAL;
	LRACTFOLLOWINGERROR : LREAL;
	XCONSTANTVELOCITY : BOOL;
	XACCELERATING : BOOL;
	XDECELERATING : BOOL;
	XDIRECTIONPOSITIVE : BOOL;
	XDIRECTIONNEGATIVE : BOOL;
END_VAR
VAR_IN_OUT
	AXIS : AXIS_REF;
END_VAR
VAR
	TM_INT : _TM_BasicMotionBase;
	PPAR : POINTER TO L_TT1P_scPar_BasicMotionBase;
	PPAR_INT : POINTER TO L_TT1P_scPar_BasicMotionBase;
	SCSIGNALFLOW : _scSF_TM_MotionControl;
	SCACCESSPOINTS : _scAP_TM_MotionControl;
END_VAR
END_FUNCTION_BLOCK

(* ---- L_TT1P_CALCPRODUCTERROR_ADVANCED.fb ---- *)
FUNCTION_BLOCK L_TT1P_CALCPRODUCTERROR_ADVANCED
VAR_INPUT
	XPRODUCTDETECTED : BOOL;
	LRACTPRODUCTPOS : LREAL;
	XENABLEPITCHCHECKING : BOOL;
	LRPRODUCTTARGET : LREAL;
	LRFACTORCOMPAREPOSITION : LREAL;
	BYNUMBEROFTARGETS : BYTE;
END_VAR
VAR_OUTPUT
	LRMASTERPOSITIONATDETECTION : LREAL;
	LRPRODUCTERROR : LREAL;
END_VAR
VAR_IN_OUT
	AXISMASTER : AXIS_REF;
END_VAR
VAR
	LRCORRECTEDFACTORCOMPAREPOSITION : LREAL;
	BCURRENTPITCH : BOOL;
	L_T01S_POSTRANSITION1 : L_TT1P_PosTransition;
	L_T01S_POSTRANSITION2 : L_TT1P_PosTransition;
	L_T01S_POSTRANSITION3 : L_TT1P_PosTransition;
	BDOUBLEPITCHCHECKACTIVE : BOOL;
	BYTARGETPITCHCHECK : BYTE;
	BYTARGETPITCHCHECKSAVED : BYTE;
	LRPRODUCTERROR1 : LREAL;
	LRPRODUCTERROR2 : LREAL;
	LRPRODUCTERROR3 : LREAL;
	LRPRODUCTTARGET1CORRECTED : LREAL;
	LRPRODUCTTARGET2CORRECTED : LREAL;
	LRPRODUCTTARGET3CORRECTED : LREAL;
	BTEST : BOOL;
	LRPRODUCTERRORFISRSTANDSECOND : LREAL;
END_VAR
END_FUNCTION_BLOCK

(* ---- L_TT1P_CALCULATEPARKPOSITION.fb ---- *)
FUNCTION_BLOCK L_TT1P_CALCULATEPARKPOSITION
VAR_INPUT
	XENABLE : BOOL;
	XEXECUTEPARKPOS : BOOL;
	LRSLAVEPOS : LREAL;
	LRPARKPOS : LREAL;
	EMODE : WORD;
END_VAR
VAR_OUTPUT
	LRPARKDISTANCE : LREAL;
END_VAR
VAR
	XEXECUTEPARKPOS_OLD : BOOL;
END_VAR
END_FUNCTION_BLOCK

(* ---- L_TT1P_CALCULATETARGETPOS.fb ---- *)
FUNCTION_BLOCK L_TT1P_CALCULATETARGETPOS
VAR_INPUT
	XRESET : BOOL;
	XENABLE : BOOL;
	XEXECUTENEXTCUT : BOOL;
	XEXECUTEFIRSTCUT : BOOL;
	XTPNOTVALID : BOOL;
	XEXECUTEGAP : BOOL;
	XRESUMETARGETPOS : BOOL;
	XSTARTFLYINGSAW : BOOL;
	XISHOMED : BOOL;
	LRHOMEPOSITION : LREAL;
	ETMSTATE : L_TT1P_States;
	XSYNCININSTANT : BOOL;
	XSETMATERIALCOUNTER : BOOL;
	LRMATERIALCOUNTER : LREAL;
	LRDELTAMATERIALPOS : LREAL;
	LRSLAVEPOS : LREAL;
	LRCUTTINGLENGTH : LREAL;
	LRMARKSENSORPOS : LREAL;
	LRGAP : LREAL;
	LRMARKPOSITION : LREAL;
	XLOADTOTALCUTTINGLENGTH : BOOL;
	LRLOADTOTALCUTTINGLENGTH : LREAL;
	XLOADTARGETPOS : BOOL;
	LRLOADTARGETPOS : LREAL;
	EMODE : L_TT1P_eModesFlyingSaw;
	LRVELINMASTER : LREAL;
	LRACCDIST : LREAL;
	LRACCTIME : LREAL;
	LRTASKCYCLETIME : LREAL;
	XEMPTYSTACK : BOOL;
	XSYNCHRONIZED : BOOL;
	XINPOSITION : BOOL;
END_VAR
VAR_OUTPUT
	XEXECUTEGAPOUT : BOOL;
	LRTARGETPOS : LREAL;
	LRTARGETPOS_OUT : LREAL;
	LRTOTALPRODUCTLENGTH : LREAL;
END_VAR
VAR
	R_TRIG1 : R_Trig;
	XEXECUTE_OLD : BOOL;
	LROFFSET_INT : LREAL;
	XGAPREQUESTED : BOOL;
	XENABLE_OLD : BOOL;
	LRDELTAMATERIALPOS_INT : LREAL;
	XEXECUTEGAP_OLD : BOOL;
	LRMATERIALCOUNTER_OLD : LREAL;
	XEXECUTENEXTCUT_OLD : BOOL;
	XSYNCININSTANT_OLD : BOOL;
	LRTOLERANCE : LREAL;
	EMODE_OLD : WORD;
	XSTARTFLYINGSAW_OLD : BOOL;
	XEXECUTEFIRSTCUT_OLD : BOOL;
	LRTOTALPRODUCTLENGTH_OLD : LREAL;
	XTPNOTVALID_OLD : BOOL;
	LRTARGETPOS_TEST : LREAL;
	LROFFSETOUT_INT : LREAL;
	XISHOMED_OLD : BOOL;
	ETMSTATE_OLD : L_TT1P_States;
	XSETMATERIALCOUNTER_OLD : BOOL;
	LRGAPTOTAL_INT : LREAL;
END_VAR
END_FUNCTION_BLOCK

(* ---- L_TT1P_CALCULATETPONMATERIALPOS.fb ---- *)
FUNCTION_BLOCK L_TT1P_CALCULATETPONMATERIALPOS
VAR_INPUT
	XENABLE : BOOL;
	BYTASKCYCLEDELAY : BYTE := 4;
	XMARKRECEIVE : BOOL;
	LRMARKSENSORPOS : LREAL;
	LRACTMARKPOSIN : LREAL;
	LRCYCPOSTPAXIS : LREAL;
	LRCYCVELTPAXIS : LREAL;
	LRCYCLELENGTHTPAXIS : LREAL;
	LRCYCLELENGTHTARGETAXIS : LREAL;
	LRTASKCYCLETIME : LREAL;
	XRESETMARKSTACK : BOOL;
	LRMATERIALCOUNTER : LREAL;
	LRUPPERLIMITWORKINGRANGE : LREAL;
	LRLOWERLIMITWORKINGRANGE : LREAL;
	LRFACTOR : LREAL;
	LRCOMPVELFACTOR : LREAL;
	XSCIPTONEXTPOSOUT : BOOL;
	XSYNCININSTANT : BOOL;
	XEXECUTEFIRSTCUT : BOOL;
	XNOMARKSTACK : BOOL;
END_VAR
VAR_OUTPUT
	LRTPPOSOUT : LREAL;
	XEXECUTEFIRSTCUT_OLD : BOOL;
	LRTPACTTIMESTAMP : LREAL;
	XFULL : BOOL;
	WMARKPOSITIONVALID : WORD;
	WININDEX : WORD;
	ALRMARKPOSITIONARRAY : ARRAY [0..15] OF LREAL := [0, 0, 0, 0, 0, 0, 0, 0, 0, 0, 0, 0, 0, 0, 0, 0];
	ALRTIMESTAMPARRAY : ARRAY [0..15] OF LREAL;
	XEMPTY : BOOL := TRUE;
	WOUTINDEX : WORD;
	BYREMAINMARKSTACK : BYTE := 15;
	XMARKRECEIVED : BOOL;
	XTPPOSVALID : BOOL;
	BYCOUNTEROUT : BYTE;
	XERROR : BOOL;
END_VAR
VAR
	R_TRIG1 : R_TRIG;
	LRTIMESTAMP : LREAL;
	BYTPIDLEINDEX : BYTE;
	BYTPACTINDEX : BYTE;
	ALRPOSITION : ARRAY [0..15] OF LREAL;
	BYTPPREVINDEX : BYTE;
	BYTMP : BYTE;
	XSKIPTONEXTPOS : BOOL;
	WTESTCOUNTER : WORD;
	XTEST : BOOL;
	XWAIT : BOOL;
	WCOUNTINVALIDTIMESTAMP : WORD;
	LRDISTINACTMASTER : LREAL;
	BYTEST : BYTE;
	LRMARKPOSITIONDIFF : LREAL;
	LRMARKPOSITIONDIFF2 : LREAL;
	LRPOSFIFOX : ARRAY [1..20] OF LREAL := [10(0)];
	LRPOSFIFOREG : ARRAY [1..20] OF LREAL := [10(0)];
	BYCOUNTER : BYTE := 1;
	LRSTACKDIFFERENCE : LREAL;
	LRTPDELTAINMS : LREAL;
	LRDELTAPCT : LREAL;
	LRTEMP : LREAL;
	IDIRECTION : INT;
	LRACTMARKPOSIN_OLD : LREAL;
	R_TRIG2 : R_TRIG;
	DWSTATE : DWORD;
	WSTOREDPOSVALUES : WORD;
	LRACTMARKPOSIN_INT : LREAL;
	XSYNCININSTANT_OLD : BOOL;
	XWAIT_OLD : BOOL;
	XRESETMARKSTACK_OLD : BOOL;
	BYCNT : BYTE;
	BYSTEPPER : BYTE;
	LRTPPOSOUT_INT : LREAL;
END_VAR
END_FUNCTION_BLOCK

METHOD SEARCHINSTACKNEGATIVE
END_METHOD

METHOD SEARCHINSTACKPOSITIVE
END_METHOD

(* ---- L_TT1P_CALCULATETPONMATERIALPOS_INTERN.fb ---- *)
FUNCTION_BLOCK L_TT1P_CALCULATETPONMATERIALPOS_INTERN
VAR_INPUT
	XENABLE : BOOL;
	BYTASKCYCLEDELAY : BYTE := 4;
	XMARKRECEIVE : BOOL;
	LRMARKSENSORPOS : LREAL;
	LRACTMARKPOSIN : LREAL;
	LRCYCPOSTPAXIS : LREAL;
	LRCYCVELTPAXIS : LREAL;
	LRCYCLELENGTHTPAXIS : LREAL;
	LRCYCLELENGTHTARGETAXIS : LREAL;
	LRTASKCYCLETIME : LREAL;
	XRESETMARKSTACK : BOOL;
	LRMATERIALCOUNTER : LREAL;
	LRUPPERLIMITWORKINGRANGE : LREAL;
	LRLOWERLIMITWORKINGRANGE : LREAL;
	LRFACTOR : LREAL;
	LRCOMPVELFACTOR : LREAL;
	XSCIPTONEXTPOSOUT : BOOL;
	XSYNCININSTANT : BOOL;
	XEXECUTEFIRSTCUT : BOOL;
END_VAR
VAR_OUTPUT
	LRTPPOSOUT : LREAL;
	XEXECUTEFIRSTCUT_OLD : BOOL;
	LRTPACTTIMESTAMP : LREAL;
	XFULL : BOOL;
	WMARKPOSITIONVALID : WORD;
	WININDEX : WORD;
	ALRMARKPOSITIONARRAY : ARRAY [0..15] OF LREAL := [0, 0, 0, 0, 0, 0, 0, 0, 0, 0, 0, 0, 0, 0, 0, 0];
	ALRTIMESTAMPARRAY : ARRAY [0..15] OF LREAL;
	XEMPTY : BOOL := TRUE;
	WOUTINDEX : WORD;
	BYREMAINMARKSTACK : BYTE := 15;
	XTPRECEIVED : BOOL;
	XMARKRECEIVED : BOOL;
	XTPPOSVALID : BOOL;
	BYCOUNTEROUT : BYTE;
	XERROR : BOOL;
END_VAR
VAR
	R_TRIG1 : R_TRIG;
	LRTIMESTAMP : LREAL;
	BYTPIDLEINDEX : BYTE;
	BYTPACTINDEX : BYTE;
	ALRPOSITION : ARRAY [0..15] OF LREAL;
	BYTPPREVINDEX : BYTE;
	BYTMP : BYTE;
	XSKIPTONEXTPOS : BOOL;
	WTESTCOUNTER : WORD;
	XTEST : BOOL;
	XWAIT : BOOL;
	WCOUNTINVALIDTIMESTAMP : WORD;
	LRDISTINACTMASTER : LREAL;
	BYTEST : BYTE;
	LRMARKPOSITIONDIFF : LREAL;
	LRMARKPOSITIONDIFF2 : LREAL;
	LRPOSFIFOX : ARRAY [1..20] OF LREAL := [10(0)];
	LRPOSFIFOREG : ARRAY [1..20] OF LREAL := [10(0)];
	BYCOUNTER : BYTE := 2;
	LRSTACKDIFFERENCE : LREAL;
	LRTPDELTAINMS : LREAL;
	LRDELTAPCT : LREAL;
	LRTEMP : LREAL;
	IDIRECTION : INT;
	LRACTMARKPOSIN_OLD : LREAL;
	R_TRIG2 : R_TRIG;
	DWSTATE : DWORD;
	WSTOREDPOSVALUES : WORD;
	LRACTMARKPOSIN_INT : LREAL;
	XSYNCININSTANT_OLD : BOOL;
	XWAIT_OLD : BOOL;
	XRESETMARKSTACK_OLD : BOOL;
	BYCNT : BYTE;
	BYSTEPPER : BYTE;
END_VAR
END_FUNCTION_BLOCK

METHOD SEARCHINSTACKNEGATIVE
END_METHOD

METHOD SEARCHINSTACKPOSITIVE
END_METHOD

(* ---- L_TT1P_CLUTCHVELOCITY.fb ---- *)
FUNCTION_BLOCK L_TT1P_CLUTCHVELOCITY
VAR_INPUT
	XENABLE : BOOL;
	XCLOSE : BOOL;
	XOPENINSTANT : BOOL;
	LRCYCVEL : LREAL;
	LRGROUNDVEL : LREAL;
	LRACCDECOPEN : LREAL;
	LRACCDECCLOSE : LREAL;
	LRDECSTOP : LREAL;
	LRJERK : LREAL;
END_VAR
VAR_OUTPUT
	XOPEN : BOOL;
	XACCDEC : BOOL;
	LRSETVELOUT : LREAL;
END_VAR
VAR
	HLP_CLUTCHV : L_TT1P_HlpRampGenerator;
	LRBASESPEED : LREAL;
	LRCLOSESPEED : LREAL;
	LRNUMERATOR : LREAL;
	LRDENUMERATOR : LREAL;
	XINITFLAG : BOOL;
	WSTEPCOUNTER : WORD;
	LRSETVELRAMPGENERATOR : LREAL;
	LRLOADRAMPGENDIFF : LREAL;
	XCOMPENSATEVELOCITYJUMP : BOOL;
	XCOMPENSATIONACTIVE : BOOL;
	CLUTCHV_INIT : WORD := 0;
	CLUTCHV_ENABLE : WORD := 1;
	CLUTCHV_CLOSE : WORD := 2;
	CLUTCHV_CLOSING : WORD := 3;
	CLUTCHV_CLOSE_DONE : WORD := 4;
	CLUTCHV_OPENING : WORD := 5;
	CLUTCHV_OPEN_STOP : WORD := 6;
	CLUTCHV_OPENINSTANT_DONE : WORD := 7;
	CLUTCHV_OPENINSTANT_DISABLE : WORD := 8;
	CLUTCHV_CLOSING_STOP : WORD := 9;
END_VAR
END_FUNCTION_BLOCK

METHOD CLUTCHCLOSINGTRANSITION
END_METHOD

METHOD CLUTCHOPENINGTRANSITION
END_METHOD

METHOD COMPENSATEVELOCITYJUMP
END_METHOD

METHOD OPENINSTANTTRANSITION
END_METHOD

(* ---- L_TT1P_CORRECTTARGETPOSITION.fb ---- *)
FUNCTION_BLOCK L_TT1P_CORRECTTARGETPOSITION
VAR_INPUT
	LRPRODUCTTARGET : LREAL;
	LRDISTANCETOOUTFEED : LREAL;
	LRMASTERPOSITIONPERIOD : LREAL;
	LRVELOCITYFACTOR : LREAL;
END_VAR
VAR_OUTPUT
	XERROR : BOOL;
	LRPRODUCTTARGETOUT : LREAL;
	LRPRODUCTTARGETCORRECTED : LREAL;
	LRDISTANCETOOUTFEEDCORR : LREAL;
END_VAR
END_FUNCTION_BLOCK

(* ---- L_TT1P_CROSSCUTTERBASE.fb ---- *)
FUNCTION_BLOCK L_TT1P_CROSSCUTTERBASE
VAR_INPUT
	XENABLEINTERNALCONTROL : BOOL;
	XENABLE : BOOL;
	SCCTRLABC : scCtrl_ABC;
	XRESETERROR : BOOL;
	XREGULATORON : BOOL;
	XSTOP : BOOL;
	XHALT : BOOL;
	SCPAR : L_TT1P_scPar_CrossCutterBase;
	SCACCESSPOINTS : L_TT1P_scAP_TM_CrossCutterBase;
	XJOGPOS : BOOL;
	XJOGNEG : BOOL;
	XHOMEEXECUTE : BOOL;
	XHOMEABSSWITCH : BOOL;
	XEXECUTEMOVETOPARKPOS : BOOL;
	XSYNCCROSSCUTTER : BOOL;
	XSYNCOUTINSTANT : BOOL;
	XHOLDINPARKPOS : BOOL;
	LRPRODUCTLENGTH : LREAL;
	LRSETOVERSPEEDSCALED : LREAL;
	LRSETOFFSETMASTER : LREAL;
	XTRIMPOS : BOOL;
	XTRIMNEG : BOOL;
	XRESETTRIMOFFSET : BOOL;
END_VAR
VAR_OUTPUT
	XINTERNALCONTROLACTIVE : BOOL;
	ETMSTATE : L_TT1P_States := L_TT1P_States.INIT;
	SCSTATUSABC : scStatus_ABC;
	XERROR : BOOL;
	XWARNING : BOOL;
	EERRORID : L_IE1P_Error;
	SCERRORINFO : L_TT1P_scErrorInfo;
	XAXISENABLED : BOOL;
	SCSIGNALFLOW : L_TT1P_scSF_TM_CrossCutterBase;
	XDONE : BOOL;
	XBUSY : BOOL;
	XISHOMED : BOOL;
	XINPARKPOS : BOOL;
	XSYNCHRONISED : BOOL;
	XACCDECSYNC : BOOL;
	XHOLDINPARKPOSACTIVE : BOOL;
	XCUTTINGACTIVE : BOOL;
	XCUTDONE : BOOL;
	LRACTCUTLENGTH : LREAL;
	BYSETTOOLNOOUT : BYTE;
	BYSETAREAOUT : BYTE;
	LROFFSET : LREAL;
	LROFFSETTRIM : LREAL := 0.0;
	LROFFSETTOTAL : LREAL;
	LRSETXPOSOUT : LREAL;
	LRSETXVELOUT : LREAL;
	LRSETXACCOUT : LREAL;
	LRACTSLAVEFOLLOWINGERROR : LREAL;
	LRACTSLAVEPOS : LREAL;
	LRACTSLAVEVEL : LREAL;
	LRSLAVEMAXVEL : LREAL;
	LRSLAVEMAXACC : LREAL;
END_VAR
VAR_IN_OUT
	MASTERAXIS : AXIS_REF;
	SLAVEAXIS : AXIS_REF;
END_VAR
VAR
	TM_INT : _TM_CrossCutterBase;
	PPAR : POINTER TO L_TT1P_scPar_CrossCutterBase;
	PPAR_INT : POINTER TO L_TT1P_scPar_CrossCutterBase;
END_VAR
END_FUNCTION_BLOCK

(* ---- L_TT1P_CROSSCUTTERSTATE.fb ---- *)
FUNCTION_BLOCK L_TT1P_CROSSCUTTERSTATE
VAR_INPUT
	XENABLEINTERNALCONTROL : BOOL;
	XENABLE : BOOL;
	SCCTRLABC : scCtrl_ABC;
	XRESETERROR : BOOL;
	XREGULATORON : BOOL;
	XSTOP : BOOL;
	XHALT : BOOL;
	SCPAR : L_TT1P_scPar_CrossCutterState;
	SCACCESSPOINTS : L_TT1P_scAP_TM_CrossCutterState;
	XJOGPOS : BOOL;
	XJOGNEG : BOOL;
	XHOMEEXECUTE : BOOL;
	XHOMEABSSWITCH : BOOL;
	XEXECUTEMOVETOPARKPOS : BOOL;
	XSYNCCROSSCUTTER : BOOL;
	XSYNCOUTINSTANT : BOOL;
	XHOLDINPARKPOS : BOOL;
	LRPRODUCTLENGTH : LREAL;
	LRSETOVERSPEEDSCALED : LREAL;
	LRSETOFFSETMASTER : LREAL;
	XTRIMPOS : BOOL;
	XTRIMNEG : BOOL;
	XRESETTRIMOFFSET : BOOL;
	XTEACHMARKWINDOW : BOOL;
	XMARKRECEIVE : BOOL;
	LRACTMARKPOSIN : LREAL;
	LRCYCPOSEXTENCODER : LREAL;
	XLOADREGPOS : BOOL;
	LRLOADREGPOS : LREAL;
	XGEARFACTORCORR : BOOL;
	XGEARFACTORCORRHOLD : BOOL;
END_VAR
VAR_OUTPUT
	XINTERNALCONTROLACTIVE : BOOL;
	ETMSTATE : L_TT1P_States := L_TT1P_States.INIT;
	SCSTATUSABC : scStatus_ABC;
	XERROR : BOOL;
	XWARNING : BOOL;
	EERRORID : L_IE1P_Error;
	SCERRORINFO : L_TT1P_scErrorInfo;
	XAXISENABLED : BOOL;
	SCSIGNALFLOW : L_TT1P_scSF_TM_CrossCutterState;
	XDONE : BOOL;
	XBUSY : BOOL;
	XISHOMED : BOOL;
	XINPARKPOS : BOOL;
	XSYNCHRONISED : BOOL;
	XACCDECSYNC : BOOL;
	XHOLDINPARKPOSACTIVE : BOOL;
	XCUTTINGACTIVE : BOOL;
	XCUTDONE : BOOL;
	LRACTCUTLENGTH : LREAL;
	BYSETTOOLNOOUT : BYTE;
	BYSETAREAOUT : BYTE;
	LROFFSET : LREAL;
	LROFFSETTRIM : LREAL;
	LROFFSETTOTAL : LREAL;
	LRSETXPOSOUT : LREAL;
	LRSETXVELOUT : LREAL;
	LRSETXACCOUT : LREAL;
	LRACTSLAVEFOLLOWINGERROR : LREAL;
	LRACTSLAVEPOS : LREAL;
	LRACTSLAVEVEL : LREAL;
	LRSLAVEMAXVEL : LREAL;
	LRSLAVEMAXACC : LREAL;
	XTRQCTRLACTIVE : BOOL;
	LRSETMOTORPRECTRLTRQOUT : LREAL;
	XREGISTERCTRLACTIVE : BOOL;
	XTEACHMARKWINDOWACTIVE : BOOL;
	LRSETREGPOSOUT : LREAL;
	LRMARKSENSORPOS : LREAL;
	LRREGMARKPOS : LREAL;
	LRACTMARKERROR : LREAL;
	LRACTMARKDIST : LREAL;
	XMARKRECEIVED : BOOL;
	XCORRACTIVE : BOOL;
	XCORRLIMITED : BOOL;
	XMARKWINDOWOPEN : BOOL;
	XMARKOUTOFWINDOW : BOOL;
	XMARKNOTDETECTED : BOOL;
	XMARKWINDOWTEACHED : BOOL;
	LRAVERAGEGEARFACTORCORR : LREAL;
	XGEARFACTORCORRLIMITED : BOOL;
END_VAR
VAR_IN_OUT
	MASTERAXIS : AXIS_REF;
	SLAVEAXIS : AXIS_REF;
END_VAR
VAR
	TM_INT : _TM_CrossCutterState;
	PPAR : POINTER TO L_TT1P_scPar_CrossCutterState;
	PPAR_INT : POINTER TO L_TT1P_scPar_CrossCutterState;
END_VAR
END_FUNCTION_BLOCK

(* ---- L_TT1P_ELECTRICALSHAFTPOSBASE.fb ---- *)
FUNCTION_BLOCK L_TT1P_ELECTRICALSHAFTPOSBASE
VAR_INPUT
	XENABLEINTERNALCONTROL : BOOL;
	XENABLE : BOOL;
	SCCTRLABC : scCtrl_ABC;
	XRESETERROR : BOOL;
	XREGULATORON : BOOL;
	XSTOP : BOOL;
	XHALT : BOOL;
	SCPAR : L_TT1P_scPar_ElectricalShaftPosBase;
	SCACCESSPOINTS : L_TT1P_scAP_ElectricalShaftPosBase;
	XJOGPOS : BOOL;
	XJOGNEG : BOOL;
	XHOMEEXECUTE : BOOL;
	XHOMEABSSWITCH : BOOL;
	XSYNCPOS : BOOL;
	LRSETOFFSETSLAVE : LREAL;
END_VAR
VAR_OUTPUT
	XINTERNALCONTROLACTIVE : BOOL;
	ETMSTATE : L_TT1P_States := L_TT1P_States.INIT;
	SCSTATUSABC : scStatus_ABC;
	XERROR : BOOL;
	XWARNING : BOOL;
	EERRORID : L_IE1P_Error;
	SCERRORINFO : L_TT1P_scErrorInfo;
	XAXISENABLED : BOOL;
	SCSIGNALFLOW : L_TT1P_scSF_ElectricalShaftPosBase;
	XDONE : BOOL;
	XBUSY : BOOL;
	XISHOMED : BOOL;
	LRACTVEL : LREAL;
	LRACTPOS : LREAL;
	LROFFSET : LREAL;
END_VAR
VAR_IN_OUT
	MASTERAXIS : AXIS_REF;
	SLAVEAXIS : AXIS_REF;
END_VAR
VAR
	TM_INT : _TM_ElectricalShaftPosBase;
	PPAR : POINTER TO L_TT1P_scPar_ElectricalShaftPosBase;
	PPAR_INT : POINTER TO L_TT1P_scPar_ElectricalShaftPosBase;
END_VAR
END_FUNCTION_BLOCK

(* ---- L_TT1P_ELECTRICALSHAFTPOSHIGH.fb ---- *)
FUNCTION_BLOCK L_TT1P_ELECTRICALSHAFTPOSHIGH
VAR_INPUT
	XENABLEINTERNALCONTROL : BOOL;
	XENABLE : BOOL;
	SCCTRLABC : scCtrl_ABC;
	XRESETERROR : BOOL;
	XREGULATORON : BOOL;
	XSTOP : BOOL;
	XHALT : BOOL;
	SCPAR : L_TT1P_scPar_ElectricalShaftPosHigh;
	SCACCESSPOINTS : L_TT1P_scAP_ElectricalShaftPosHigh;
	XJOGPOS : BOOL;
	XJOGNEG : BOOL;
	XHOMEEXECUTE : BOOL;
	XHOMEABSSWITCH : BOOL;
	XSYNCPOS : BOOL;
	LRSETOFFSETMASTER : LREAL;
	LRSETOFFSETSLAVE : LREAL;
	XTRIMPOS : BOOL;
	XTRIMNEG : BOOL;
	XSYNCINSTANT : BOOL;
	XSYNCOUTINSTANT : BOOL;
	XSYNCPOSRESTORE : BOOL;
END_VAR
VAR_OUTPUT
	XINTERNALCONTROLACTIVE : BOOL;
	ETMSTATE : L_TT1P_States := L_TT1P_States.INIT;
	SCSTATUSABC : scStatus_ABC;
	XERROR : BOOL;
	XWARNING : BOOL;
	EERRORID : L_IE1P_Error;
	SCERRORINFO : L_TT1P_scErrorInfo;
	XAXISENABLED : BOOL;
	SCSIGNALFLOW : L_TT1P_scSF_ElectricalShaftPosHigh;
	XDONE : BOOL;
	XBUSY : BOOL;
	XISHOMED : BOOL;
	LRACTVEL : LREAL;
	LRACTPOS : LREAL;
	LROFFSET : LREAL;
	LROFFSETTRIM : LREAL;
	LROFFSETTOTAL : LREAL;
	XSYNCHRONISED : BOOL;
	XACCDECSYNC : BOOL;
	LROFFSETSYNCPOS : LREAL;
	LROFFSETMASTER : LREAL;
END_VAR
VAR_IN_OUT
	MASTERAXIS : AXIS_REF;
	SLAVEAXIS : AXIS_REF;
END_VAR
VAR
	TM_INT : _TM_ElectricalShaftPosHigh;
	PPAR : POINTER TO L_TT1P_scPar_ElectricalShaftPosHigh;
	PPAR_INT : POINTER TO L_TT1P_scPar_ElectricalShaftPosHigh;
END_VAR
END_FUNCTION_BLOCK

(* ---- L_TT1P_ELECTRICALSHAFTPOSSTATE.fb ---- *)
FUNCTION_BLOCK L_TT1P_ELECTRICALSHAFTPOSSTATE
VAR_INPUT
	XENABLEINTERNALCONTROL : BOOL;
	XENABLE : BOOL;
	SCCTRLABC : scCtrl_ABC;
	XRESETERROR : BOOL;
	XREGULATORON : BOOL;
	XSTOP : BOOL;
	XHALT : BOOL;
	SCPAR : L_TT1P_scPar_ElectricalShaftPosState;
	SCACCESSPOINTS : L_TT1P_scAP_ElectricalShaftPosState;
	XJOGPOS : BOOL;
	XJOGNEG : BOOL;
	XHOMEEXECUTE : BOOL;
	XHOMEABSSWITCH : BOOL;
	XSYNCPOS : BOOL;
	LRSETOFFSETSLAVE : LREAL;
	XTRIMPOS : BOOL;
	XTRIMNEG : BOOL;
END_VAR
VAR_OUTPUT
	XINTERNALCONTROLACTIVE : BOOL;
	ETMSTATE : L_TT1P_States := L_TT1P_States.INIT;
	SCSTATUSABC : scStatus_ABC;
	XERROR : BOOL;
	XWARNING : BOOL;
	EERRORID : L_IE1P_Error;
	SCERRORINFO : L_TT1P_scErrorInfo;
	XAXISENABLED : BOOL;
	SCSIGNALFLOW : L_TT1P_scSF_ElectricalShaftPosState;
	XDONE : BOOL;
	XBUSY : BOOL;
	XISHOMED : BOOL;
	LRACTVEL : LREAL;
	LRACTPOS : LREAL;
	LROFFSET : LREAL;
	LROFFSETTRIM : LREAL;
	LROFFSETTOTAL : LREAL;
	XSYNCHRONISED : BOOL;
	XACCDECSYNC : BOOL;
END_VAR
VAR_IN_OUT
	MASTERAXIS : AXIS_REF;
	SLAVEAXIS : AXIS_REF;
END_VAR
VAR
	TM_INT : _TM_ElectricalShaftPosState;
	PPAR : POINTER TO L_TT1P_scPar_ElectricalShaftPosState;
	PPAR_INT : POINTER TO L_TT1P_scPar_ElectricalShaftPosState;
END_VAR
END_FUNCTION_BLOCK

(* ---- L_TT1P_ELECTRICALSHAFTVELBASE.fb ---- *)
FUNCTION_BLOCK L_TT1P_ELECTRICALSHAFTVELBASE
VAR_INPUT
	XENABLEINTERNALCONTROL : BOOL;
	XENABLE : BOOL;
	SCCTRLABC : scCtrl_ABC;
	XRESETERROR : BOOL;
	XREGULATORON : BOOL;
	XSTOP : BOOL;
	XHALT : BOOL;
	SCPAR : L_TT1P_scPar_ElectricalShaftVelBase;
	SCACCESSPOINTS : L_TT1P_scAP_ElectricalShaftVelBase;
	XJOGPOS : BOOL;
	XJOGNEG : BOOL;
	XSYNCVEL : BOOL;
	LRSETOFFSET : LREAL;
END_VAR
VAR_OUTPUT
	XINTERNALCONTROLACTIVE : BOOL;
	ETMSTATE : L_TT1P_States := L_TT1P_States.INIT;
	SCSTATUSABC : scStatus_ABC;
	XERROR : BOOL;
	XWARNING : BOOL;
	EERRORID : L_IE1P_Error;
	SCERRORINFO : L_TT1P_scErrorInfo;
	XAXISENABLED : BOOL;
	SCSIGNALFLOW : L_TT1P_scSF_ElectricalShaftVelBase;
	XDONE : BOOL;
	XBUSY : BOOL;
	LRACTVEL : LREAL;
	LRACTPOS : LREAL;
	LROFFSET : LREAL;
END_VAR
VAR_IN_OUT
	MASTERAXIS : AXIS_REF;
	SLAVEAXIS : AXIS_REF;
END_VAR
VAR
	TM_INT : _TM_ElectricalShaftVelBase;
	PPAR : POINTER TO L_TT1P_scPar_ElectricalShaftVelBase;
	PPAR_INT : POINTER TO L_TT1P_scPar_ElectricalShaftVelBase;
	XHOMEEXECUTE : BOOL;
	XHOMEABSSWITCH : BOOL;
	XISHOMED : BOOL;
END_VAR
END_FUNCTION_BLOCK

(* ---- L_TT1P_ELECTRICALSHAFTVELHIGH.fb ---- *)
FUNCTION_BLOCK L_TT1P_ELECTRICALSHAFTVELHIGH
VAR_INPUT
	XENABLEINTERNALCONTROL : BOOL;
	XENABLE : BOOL;
	SCCTRLABC : scCtrl_ABC;
	XRESETERROR : BOOL;
	XREGULATORON : BOOL;
	XSTOP : BOOL;
	XHALT : BOOL;
	SCPAR : L_TT1P_scPar_ElectricalShaftVelHigh;
	SCACCESSPOINTS : L_TT1P_scAP_ElectricalShaftVelHigh;
	XJOGPOS : BOOL;
	XJOGNEG : BOOL;
	XSYNCVEL : BOOL;
	LRSETOFFSET : LREAL;
	XTRIMPOS : BOOL;
	XTRIMNEG : BOOL;
	LRSETGROUNDVEL : LREAL;
END_VAR
VAR_OUTPUT
	XINTERNALCONTROLACTIVE : BOOL;
	ETMSTATE : L_TT1P_States := L_TT1P_States.INIT;
	SCSTATUSABC : scStatus_ABC;
	XERROR : BOOL;
	XWARNING : BOOL;
	EERRORID : L_IE1P_Error;
	SCERRORINFO : L_TT1P_scErrorInfo;
	XAXISENABLED : BOOL;
	SCSIGNALFLOW : L_TT1P_scSF_ElectricalShaftVelHigh;
	XDONE : BOOL;
	XBUSY : BOOL;
	LRACTVEL : LREAL;
	LRACTPOS : LREAL;
	LROFFSET : LREAL;
	LROFFSETTRIM : LREAL;
	LROFFSETTOTAL : LREAL;
	XSYNCHRONISED : BOOL;
	XACCDECSYNC : BOOL;
END_VAR
VAR_IN_OUT
	MASTERAXIS : AXIS_REF;
	SLAVEAXIS : AXIS_REF;
END_VAR
VAR
	TM_INT : _TM_ElectricalShaftVelHigh;
	PPAR : POINTER TO L_TT1P_scPar_ElectricalShaftVelHigh;
	PPAR_INT : POINTER TO L_TT1P_scPar_ElectricalShaftVelHigh;
	XHOMEEXECUTE : BOOL;
	XHOMEABSSWITCH : BOOL;
	XISHOMED : BOOL;
END_VAR
END_FUNCTION_BLOCK

(* ---- L_TT1P_ELECTRICALSHAFTVELSTATE.fb ---- *)
FUNCTION_BLOCK L_TT1P_ELECTRICALSHAFTVELSTATE
VAR_INPUT
	XENABLEINTERNALCONTROL : BOOL;
	XENABLE : BOOL;
	SCCTRLABC : scCtrl_ABC;
	XRESETERROR : BOOL;
	XREGULATORON : BOOL;
	XSTOP : BOOL;
	XHALT : BOOL;
	SCPAR : L_TT1P_scPar_ElectricalShaftVelState;
	SCACCESSPOINTS : L_TT1P_scAP_ElectricalShaftVelState;
	XJOGPOS : BOOL;
	XJOGNEG : BOOL;
	XSYNCVEL : BOOL;
	LRSETOFFSET : LREAL;
	XTRIMPOS : BOOL;
	XTRIMNEG : BOOL;
END_VAR
VAR_OUTPUT
	XINTERNALCONTROLACTIVE : BOOL;
	ETMSTATE : L_TT1P_States := L_TT1P_States.INIT;
	SCSTATUSABC : scStatus_ABC;
	XERROR : BOOL;
	XWARNING : BOOL;
	EERRORID : L_IE1P_Error;
	SCERRORINFO : L_TT1P_scErrorInfo;
	XAXISENABLED : BOOL;
	SCSIGNALFLOW : L_TT1P_scSF_ElectricalShaftVelState;
	XDONE : BOOL;
	XBUSY : BOOL;
	LRACTVEL : LREAL;
	LRACTPOS : LREAL;
	LROFFSET : LREAL;
	LROFFSETTRIM : LREAL;
	LROFFSETTOTAL : LREAL;
	XSYNCHRONISED : BOOL;
	XACCDECSYNC : BOOL;
END_VAR
VAR_IN_OUT
	MASTERAXIS : AXIS_REF;
	SLAVEAXIS : AXIS_REF;
END_VAR
VAR
	TM_INT : _TM_ElectricalShaftVelState;
	PPAR : POINTER TO L_TT1P_scPar_ElectricalShaftVelState;
	PPAR_INT : POINTER TO L_TT1P_scPar_ElectricalShaftVelState;
	XHOMEEXECUTE : BOOL;
	XHOMEABSSWITCH : BOOL;
	XISHOMED : BOOL;
END_VAR
END_FUNCTION_BLOCK

(* ---- L_TT1P_FILTERPRODUCTDETECTION.fb ---- *)
FUNCTION_BLOCK L_TT1P_FILTERPRODUCTDETECTION
VAR_INPUT
	XPRODUCTTRIGGERRISE : BOOL;
	XPRODUCTTRIGGERFALL : BOOL;
	LRLASTSCANOUT : LREAL;
	LRFILTERDISTPRODDETECTIONRISINGEDGE : LREAL;
	LRFILTERDISTPRODDETECTIONFALLINGEDGE : LREAL;
END_VAR
VAR_OUTPUT
	XPRODUCTDETECTED : BOOL;
	LRFILTERDISTINTEGRATOR : LREAL;
END_VAR
VAR_IN_OUT
	AXISSMARTTRACK : AXIS_REF;
END_VAR
VAR
	LRDELTAPOSITION : LREAL;
	BYSTEPPER : BYTE;
END_VAR
END_FUNCTION_BLOCK

(* ---- L_TT1P_FLEXCAMBASE.fb ---- *)
FUNCTION_BLOCK L_TT1P_FLEXCAMBASE
VAR_INPUT
	XENABLEINTERNALCONTROL : BOOL;
	XENABLE : BOOL;
	SCCTRLABC : scCtrl_ABC;
	XRESETERROR : BOOL;
	XREGULATORON : BOOL;
	XSTOP : BOOL;
	XHALT : BOOL;
	SCPAR : L_TT1P_scPar_FlexCamBase;
	SCACCESSPOINTS : L_TT1P_scAP_FlexCamBase;
	XJOGPOS : BOOL;
	XJOGNEG : BOOL;
	XHOMEEXECUTE : BOOL;
	XHOMEABSSWITCH : BOOL;
	XENABLEHWLIMIT : BOOL;
	XHWLIMITPOS : BOOL;
	XHWLIMITNEG : BOOL;
	XSYNCCAM : BOOL;
	XSYNCOUTINSTANT : BOOL;
	XCAMCHANGEINSTANT : BOOL;
	LRSETOFFSETMASTER : LREAL;
	LRSETOFFSETSLAVE : LREAL;
	LRSETSCALINGMASTER : LREAL;
	LRSETSCALINGSLAVE : LREAL;
	CAMTABLE1 : MC_CAM_REF;
END_VAR
VAR_OUTPUT
	XINTERNALCONTROLACTIVE : BOOL;
	ETMSTATE : L_TT1P_States;
	SCSTATUSABC : scStatus_ABC;
	XERROR : BOOL;
	XWARNING : BOOL;
	EERRORID : L_IE1P_Error;
	SCERRORINFO : L_TT1P_scErrorInfo;
	XAXISENABLED : BOOL;
	SCSIGNALFLOW : L_TT1P_scSF_FlexCamBase;
	XDONE : BOOL;
	XBUSY : BOOL;
	XISHOMED : BOOL;
	XHWLIMITSWITCHNEG : BOOL;
	XHWLIMITSWITCHPOS : BOOL;
	XSWLIMITENABLED : BOOL;
	XSWLIMITSWITCHACTIVE : BOOL;
	XCAMSYNCHRONISED : BOOL;
	XACCDECSYNC : BOOL;
	XENDOFPROFILE : BOOL;
	LRSETXPOSOUT : LREAL;
	LRSETXVELOUT : LREAL;
	LRSETXACCOUT : LREAL;
	LRSETYPOSOUT : LREAL;
	LRSETYVELOUT : LREAL;
	LRSETYACCOUT : LREAL;
	LRACTSLAVEPOS : LREAL;
	LRACTSLAVEVEL : LREAL;
	LRSETOFFSETMASTEROUT : LREAL;
	LRSETOFFSETSLAVEOUT : LREAL;
	LRSLAVEMAXPOS : LREAL;
	LRSLAVEMINPOS : LREAL;
	LRSLAVEMAXVEL : LREAL;
	LRSLAVEMAXACC : LREAL;
END_VAR
VAR_IN_OUT
	MASTERAXIS : AXIS_REF;
	SLAVEAXIS : AXIS_REF;
END_VAR
VAR
	TM_INT : _TM_FlexCamBaseExtension;
	PPAR : POINTER TO L_TT1P_scPar_FlexCamBase;
	PPAR_INT : POINTER TO L_TT1P_scPar_FlexCamBase;
END_VAR
END_FUNCTION_BLOCK

METHOD GET_INTERNCAMTABLE : MC_CAM_REF
END_METHOD

METHOD GET_LRCAMXEND : LREAL
END_METHOD

METHOD GET_LRCAMXSTART : LREAL
END_METHOD

METHOD GET_LRCAMYEND : LREAL
END_METHOD

METHOD GET_LRCAMYSTART : LREAL
END_METHOD

METHOD GET_STCAMNAME : STRING
END_METHOD

METHOD GET_XCOMMUNICATION : BOOL
END_METHOD

(* ---- L_TT1P_FLEXCAMSTATE.fb ---- *)
FUNCTION_BLOCK L_TT1P_FLEXCAMSTATE
VAR_INPUT
	XENABLEINTERNALCONTROL : BOOL;
	XENABLE : BOOL;
	SCCTRLABC : scCtrl_ABC;
	XRESETERROR : BOOL;
	XREGULATORON : BOOL;
	XSTOP : BOOL;
	XHALT : BOOL;
	SCPAR : L_TT1P_scPar_FlexCamState;
	SCACCESSPOINTS : L_TT1P_scAP_FlexCamState;
	XJOGPOS : BOOL;
	XJOGNEG : BOOL;
	XHOMEEXECUTE : BOOL;
	XHOMEABSSWITCH : BOOL;
	XENABLEHWLIMIT : BOOL;
	XHWLIMITPOS : BOOL;
	XHWLIMITNEG : BOOL;
	XSYNCCAM : BOOL;
	XSYNCOUTINSTANT : BOOL;
	XCAMCHANGEINSTANT : BOOL;
	LRSETOFFSETMASTER : LREAL;
	LRSETOFFSETSLAVE : LREAL;
	LRSETSCALINGMASTER : LREAL;
	LRSETSCALINGSLAVE : LREAL;
	CAMTABLE1 : MC_CAM_REF;
	CAMTABLE2 : MC_CAM_REF;
	CAMTABLE3 : MC_CAM_REF;
	CAMTABLE4 : MC_CAM_REF;
	ESETCAMTABLE : L_TT1P_CamTable := 1;
	XCAMSEQUENCER : BOOL;
END_VAR
VAR_OUTPUT
	XINTERNALCONTROLACTIVE : BOOL;
	ETMSTATE : L_TT1P_States;
	SCSTATUSABC : scStatus_ABC;
	XERROR : BOOL;
	XWARNING : BOOL;
	EERRORID : L_IE1P_Error;
	SCERRORINFO : L_TT1P_scErrorInfo;
	XAXISENABLED : BOOL;
	SCSIGNALFLOW : L_TT1P_scSF_FlexCamState;
	XDONE : BOOL;
	XBUSY : BOOL;
	XISHOMED : BOOL;
	XHWLIMITSWITCHNEG : BOOL;
	XHWLIMITSWITCHPOS : BOOL;
	XSWLIMITENABLED : BOOL;
	XSWLIMITSWITCHACTIVE : BOOL;
	XCAMSYNCHRONISED : BOOL;
	XACCDECSYNC : BOOL;
	XENDOFPROFILE : BOOL;
	LRSETXPOSOUT : LREAL;
	LRSETXVELOUT : LREAL;
	LRSETXACCOUT : LREAL;
	LRSETYPOSOUT : LREAL;
	LRSETYVELOUT : LREAL;
	LRSETYACCOUT : LREAL;
	LRACTSLAVEPOS : LREAL;
	LRACTSLAVEVEL : LREAL;
	LRSETOFFSETMASTEROUT : LREAL;
	LRSETOFFSETSLAVEOUT : LREAL;
	LRSLAVEMAXPOS : LREAL;
	LRSLAVEMINPOS : LREAL;
	LRSLAVEMAXVEL : LREAL;
	LRSLAVEMAXACC : LREAL;
	ESETCAMTABLEOUT : L_TT1P_CamTable;
	XCAMSEQUENCERACTIVE : BOOL;
END_VAR
VAR_IN_OUT
	MASTERAXIS : AXIS_REF;
	SLAVEAXIS : AXIS_REF;
END_VAR
VAR
	TM_INT : _TM_FlexCamState;
	PPAR : POINTER TO L_TT1P_scPar_FlexCamState;
	PPAR_INT : POINTER TO L_TT1P_scPar_FlexCamState;
END_VAR
END_FUNCTION_BLOCK

METHOD GET_INTERNCAMTABLE : MC_CAM_REF
END_METHOD

METHOD GET_LRCAMXEND : LREAL
END_METHOD

METHOD GET_LRCAMXSTART : LREAL
END_METHOD

METHOD GET_LRCAMYEND : LREAL
END_METHOD

METHOD GET_LRCAMYSTART : LREAL
END_METHOD

METHOD GET_STCAMNAME : STRING
END_METHOD

METHOD GET_XCOMMUNICATION : BOOL
END_METHOD

(* ---- L_TT1P_FLYINGSAWBASE.fb ---- *)
FUNCTION_BLOCK L_TT1P_FLYINGSAWBASE
VAR_INPUT
	XENABLEINTERNALCONTROL : BOOL;
	XENABLE : BOOL;
	SCCTRLABC : scCtrl_ABC;
	XRESETERROR : BOOL;
	XREGULATORON : BOOL;
	XSTOP : BOOL;
	XHALT : BOOL;
	SCPAR : L_TT1P_scPar_FlyingSawBase;
	SCACCESSPOINTS : L_TT1P_scAP_FlyingSawBase;
	XJOGPOS : BOOL;
	XJOGNEG : BOOL;
	XHOMEEXECUTE : BOOL;
	XHOMEABSSWITCH : BOOL;
	XENABLEHWLIMIT : BOOL;
	XHWLIMITPOS : BOOL;
	XHWLIMITNEG : BOOL;
	XSTARTFLYINGSAW : BOOL;
	XSYNCININSTANT : BOOL;
	XEXECUTENEXTCUT : BOOL;
	XEXECUTEGAP : BOOL;
	LRCUTTINGLENGTH : LREAL;
	XSETMATERIALCOUNTER : BOOL;
END_VAR
VAR_OUTPUT
	XINTERNALCONTROLACTIVE : BOOL;
	ETMSTATE : L_TT1P_States := L_TT1P_States.INIT;
	SCSTATUSABC : scStatus_ABC;
	XERROR : BOOL;
	XWARNING : BOOL;
	EERRORID : L_IE1P_Error;
	SCERRORINFO : L_TT1P_scErrorInfo;
	XAXISENABLED : BOOL;
	SCSIGNALFLOW : L_TT1P_scSF_FlyingSawBase;
	XDONE : BOOL;
	XBUSY : BOOL;
	XISHOMED : BOOL;
	XHWLIMITSWITCHNEG : BOOL;
	XHWLIMITSWITCHPOS : BOOL;
	XSWLIMITENABLED : BOOL;
	XSWLIMITSWITCHACTIVE : BOOL;
	XSYNCHRONISED : BOOL;
	XACCDECSYNC : BOOL;
	XINPOSITION : BOOL;
	XPOSITIONING : BOOL;
	LRACTPOS : LREAL;
	LRACTVEL : LREAL;
	LRACTFOLLOWINGERROR : LREAL;
	LRMATERIALCOUNTER : LREAL;
	LRTARGETPOS : LREAL;
	LRCUTGAP : LREAL;
END_VAR
VAR_IN_OUT
	MASTERAXIS : AXIS_REF;
	SLAVEAXIS : AXIS_REF;
END_VAR
VAR
	TM_INT : _TM_FlyingSawBase;
	PPAR : POINTER TO L_TT1P_scPar_FlyingSawBase;
	PPAR_INT : POINTER TO L_TT1P_scPar_FlyingSawBase;
END_VAR
END_FUNCTION_BLOCK

(* ---- L_TT1P_FLYINGSAWSTATE.fb ---- *)
FUNCTION_BLOCK L_TT1P_FLYINGSAWSTATE
VAR_INPUT
	XENABLEINTERNALCONTROL : BOOL;
	XENABLE : BOOL;
	SCCTRLABC : scCtrl_ABC;
	XRESETERROR : BOOL;
	XREGULATORON : BOOL;
	XSTOP : BOOL;
	XHALT : BOOL;
	SCPAR : L_TT1P_scPar_FlyingSawState;
	SCACCESSPOINTS : L_TT1P_scAP_FlyingSawState;
	XJOGPOS : BOOL;
	XJOGNEG : BOOL;
	XHOMEEXECUTE : BOOL;
	XHOMEABSSWITCH : BOOL;
	XENABLEHWLIMIT : BOOL;
	XHWLIMITPOS : BOOL;
	XHWLIMITNEG : BOOL;
	XSTARTFLYINGSAW : BOOL;
	XSYNCININSTANT : BOOL;
	XEXECUTENEXTCUT : BOOL;
	XEXECUTEGAP : BOOL;
	LRCUTTINGLENGTH : LREAL;
	XSETMATERIALCOUNTER : BOOL;
	XMOVETOPARKPOS : BOOL;
	XRESUMETARGETPOS : BOOL;
	XRESETMARKSTACK : BOOL;
	XMARKRECEIVE : BOOL;
	LRACTMARKPOSIN : LREAL;
END_VAR
VAR_OUTPUT
	XINTERNALCONTROLACTIVE : BOOL;
	ETMSTATE : L_TT1P_States := L_TT1P_States.INIT;
	SCSTATUSABC : scStatus_ABC;
	XERROR : BOOL;
	XWARNING : BOOL;
	EERRORID : L_IE1P_Error;
	SCERRORINFO : L_TT1P_scErrorInfo;
	XAXISENABLED : BOOL;
	SCSIGNALFLOW : L_TT1P_scSF_FlyingSawState;
	XDONE : BOOL;
	XBUSY : BOOL;
	XISHOMED : BOOL;
	XHWLIMITSWITCHNEG : BOOL;
	XHWLIMITSWITCHPOS : BOOL;
	XSWLIMITENABLED : BOOL;
	XSWLIMITSWITCHACTIVE : BOOL;
	XSYNCHRONISED : BOOL;
	XACCDECSYNC : BOOL;
	XINPOSITION : BOOL;
	XPOSITIONING : BOOL;
	LRACTPOS : LREAL;
	LRACTVEL : LREAL;
	LRACTFOLLOWINGERROR : LREAL;
	LRMATERIALCOUNTER : LREAL;
	LRTARGETPOS : LREAL;
	LRCUTGAP : LREAL;
	BYREMAINMARKSTACK : BYTE;
END_VAR
VAR_IN_OUT
	MASTERAXIS : AXIS_REF;
	SLAVEAXIS : AXIS_REF;
END_VAR
VAR
	TM_INT : _TM_FlyingSawState;
	PPAR : POINTER TO L_TT1P_scPar_FlyingSawState;
	PPAR_INT : POINTER TO L_TT1P_scPar_FlyingSawState;
END_VAR
END_FUNCTION_BLOCK

(* ---- L_TT1P_HLPRAMPGENERATOR.fb ---- *)
FUNCTION_BLOCK L_TT1P_HLPRAMPGENERATOR
VAR_INPUT
	LRACC : LREAL;
	LRDEC : LREAL;
	LRVEL : LREAL;
	LRJERKACC : LREAL;
	LRJERKDEC : LREAL;
	LRTASKCYCLE : LREAL;
END_VAR
VAR_OUTPUT
	LRSETVEL : LREAL;
	LRSETACCDEC : LREAL;
	DNSTATE : DINT;
END_VAR
VAR
	ALRACCLIMIT : ARRAY [0..1] OF LREAL;
	ALRJERKABS : ARRAY [0..1] OF LREAL;
	LRVELINTERNAL : LREAL;
	DWINDEX : DWORD;
	LRVELDIFF : LREAL;
	LRVELCOMPARE : LREAL;
	LRACCINTERNAL : LREAL;
	C_RG_ACC : WORD := 0;
	C_RG_DEC : WORD := 1;
	C_RG_MINJERK : LREAL := 1;
	C_RG_STATE_INI : DINT := 0;
	C_RG_STATE_CNS : DINT := 1;
	C_RG_STATE_ACC : DINT := 2;
	C_RG_STATE_DEC : DINT := 3;
END_VAR
END_FUNCTION_BLOCK

METHOD RG_GETDEC : BOOL
VAR_INPUT
	LRVELDIFF : LREAL;
	LRVEL : LREAL;
END_VAR
END_METHOD

METHOD RG_MAXJERKINDEX : WORD
VAR_INPUT
	VAR1 : LREAL;
	VAR2 : LREAL;
	IND1 : WORD;
	IND2 : WORD;
END_VAR
END_METHOD

METHOD RG_REDACC : BOOL
VAR_INPUT
	LRVELDIFF : LREAL;
	LRACC : LREAL;
END_VAR
END_METHOD

METHOD SETSTARTVALUES
VAR_INPUT
	LRVEL : LREAL;
	LRACC : LREAL;
END_VAR
END_METHOD

METHOD TFM_RG_CALCDELTAVEL
END_METHOD

METHOD TFM_RG_CALCJERK : LREAL
VAR_INPUT
	VEL : LREAL;
	ACC : LREAL;
END_VAR
END_METHOD

METHOD TFM_RG_CALCPARAMETER
END_METHOD

METHOD TFM_RG_REDACC
END_METHOD

METHOD TFM_RG_VELDIFFNEG
END_METHOD

METHOD TFM_RG_VELDIFFPOS
END_METHOD

METHOD TFM_RG_VELTARGET
END_METHOD

(* ---- L_TT1P_INPOSITION.fb ---- *)
FUNCTION_BLOCK L_TT1P_INPOSITION
VAR_INPUT
	XENABLE : BOOL;
	LRPOSWINDOW : LREAL;
	LRPOSTIME : LREAL;
	XHOLDSETPOS : BOOL;
END_VAR
VAR_OUTPUT
	XINPOSITION : BOOL;
	XBUSY : BOOL;
	LRHOLDPOSITION : LREAL;
	XERROR : BOOL;
	EERRORID : L_IE1P_Error;
END_VAR
VAR_IN_OUT
	AXIS : AXIS_REF;
END_VAR
VAR
	XINTOL : BOOL;
	XENABLEOLD : BOOL := FALSE;
	XHOLDSETPOSOLD : BOOL := FALSE;
	LRSETPOSITIONOLD : LREAL;
	XSETPOSITIONCHG : BOOL;
	INPOSITION_TON : TON;
	INPOSITION_F_TRIG : F_TRIG;
	TIMEOUT_TON : TON;
END_VAR
END_FUNCTION_BLOCK

METHOD FB_RESET : BOOL
END_METHOD

(* ---- L_TT1P_LIMITPRODUCTERROR.fb ---- *)
FUNCTION_BLOCK L_TT1P_LIMITPRODUCTERROR
VAR_INPUT
	LRPRODUCTERROR : LREAL;
	LRMAXIMUMERRORPOSITIVE : LREAL := 100;
	LRMAXIMUMERRORNEGATIVE : LREAL := 100;
END_VAR
VAR_OUTPUT
	LRPRODUCTERRORLIMITED : LREAL;
	XPRODUCTERRORLIMITED : BOOL;
END_VAR
END_FUNCTION_BLOCK

(* ---- L_TT1P_PICKANDPLACEBASE.fb ---- *)
FUNCTION_BLOCK L_TT1P_PICKANDPLACEBASE
VAR_INPUT
	XENABLEINTERNALCONTROL : BOOL;
	XENABLE : BOOL;
	SCCTRLAGBC : scCtrl_AGBC;
	XRESETERROR : BOOL;
	XREGULATORONALL : BOOL;
	XPATHSTOP : BOOL;
	XPATHHALT : BOOL;
	XSTOPALL : BOOL;
	SCPAR : L_TT1P_scPar_PickAndPlaceBase;
	SCACCESSPOINTS : L_TT1P_scAP_PickAndPlaceBase;
	XEXECUTEPICKANDPLACE : BOOL;
	XPATHINTERRUPT : BOOL;
	XGROUPHOMEEXECUTE : BOOL;
	AXHOMEABSSWITCH : ARRAY [1..12] OF BOOL;
	XGROUPENABLEHWLIMIT : BOOL;
	AXHWLIMITPOS : ARRAY [1..18] OF BOOL;
	AXHWLIMITNEG : ARRAY [1..18] OF BOOL;
	ESELECTAXIS : IDENT_IN_GROUP_REF;
	XJOGPOS : BOOL;
	XJOGNEG : BOOL;
	XABORT : BOOL;
	LROVERRIDE : LREAL := 1;
END_VAR
VAR_OUTPUT
	XINTERNALCONTROLACTIVE : BOOL;
	ETMSTATE : L_TT1P_States := L_TT1P_States.INIT;
	SCSTATUSAGBC : scStatus_AGBC;
	XERROR : BOOL;
	XWARNING : BOOL;
	EERRORID : L_IE1P_Error;
	ASCERRORINFO : ARRAY [1..18] OF L_TT1P_scErrorInfo;
	XAXESENABLED : BOOL;
	XAXESGROUPENABLED : BOOL;
	SCSIGNALFLOW : L_TT1P_scSF_PickAndPlaceBase;
	XDONE : BOOL;
	XBUSY : BOOL;
	XACTIVE : BOOL;
	XAXESGROUPHOMED : BOOL;
	XINPOSITION : BOOL;
	XHWLIMITSWITCHACTIVE : BOOL;
	XSWLIMITSWITCHACTIVE : BOOL;
	AXHWLIMITSWITCHNEG : ARRAY [1..18] OF BOOL;
	AXHWLIMITSWITCHPOS : ARRAY [1..18] OF BOOL;
	AXSWLIMITSWITCHENABLE : ARRAY [1..18] OF BOOL;
	AXSWLIMITSWITCHACTIVE : ARRAY [1..18] OF BOOL;
	XPATHHOLD : BOOL;
	XGRIPPERCTRLACTIVE : BOOL;
	XPULSEGRIPPER : BOOL;
	LRSETPATHVELOUT : LREAL;
	LRPATHPREPARATIONTIME : LREAL;
	LRPRECALCPROFILETIME : LREAL;
	ALRACTAXISPOS : ARRAY [1..18] OF LREAL;
	ALRACTAXISVEL : ARRAY [1..18] OF LREAL;
	IPROFILEPOINTPASSED : INT;
END_VAR
VAR_IN_OUT
	AXESGROUP : AXES_GROUP_KIN;
END_VAR
VAR
	TM_INT : _TM_PickAndPlaceBaseExtension;
	PPAR : POINTER TO L_TT1P_scPar_PickAndPlaceBase;
	PPAR_INT : POINTER TO L_TT1P_scPar_PickAndPlaceBase;
	FB_LIMITDYNAMICSMAINAXES : L_MC4P_LimitDynamicsMainAxes;
	FB_LIMITDYNAMICSAUXAXES : L_MC4P_LimitDynamicsAuxAxes;
	AFB_HWLIMITAXIS : ARRAY [1..13] OF L_MC1P_HWLimitSwitchInterface;
END_VAR
END_FUNCTION_BLOCK

(* ---- L_TT1P_PICKANDPLACEHIGH.fb ---- *)
FUNCTION_BLOCK L_TT1P_PICKANDPLACEHIGH
VAR_INPUT
	XENABLEINTERNALCONTROL : BOOL;
	XENABLE : BOOL;
	SCCTRLAGBC : scCtrl_AGBC;
	XRESETERROR : BOOL;
	XREGULATORONALL : BOOL;
	XPATHSTOP : BOOL;
	XPATHHALT : BOOL;
	XSTOPALL : BOOL;
	SCPAR : L_TT1P_scPar_PickAndPlaceHigh;
	SCACCESSPOINTS : L_TT1P_scAP_PickAndPlaceHigh;
	XEXECUTEPICKANDPLACE : BOOL;
	XPATHINTERRUPT : BOOL;
	XGROUPHOMEEXECUTE : BOOL;
	AXHOMEABSSWITCH : ARRAY [1..12] OF BOOL;
	XGROUPENABLEHWLIMIT : BOOL;
	AXHWLIMITPOS : ARRAY [1..18] OF BOOL;
	AXHWLIMITNEG : ARRAY [1..18] OF BOOL;
	ESELECTAXIS : IDENT_IN_GROUP_REF;
	XJOGPOS : BOOL;
	XJOGNEG : BOOL;
	XABORT : BOOL;
	LROVERRIDE : LREAL := 1;
	XACKPATHHALT : BOOL;
	XADDPROFILE : BOOL;
END_VAR
VAR_OUTPUT
	XINTERNALCONTROLACTIVE : BOOL;
	ETMSTATE : L_TT1P_States := L_TT1P_States.INIT;
	SCSTATUSAGBC : scStatus_AGBC;
	XERROR : BOOL;
	XWARNING : BOOL;
	EERRORID : L_IE1P_Error;
	ASCERRORINFO : ARRAY [1..18] OF L_TT1P_scErrorInfo;
	XAXESENABLED : BOOL;
	XAXESGROUPENABLED : BOOL;
	SCSIGNALFLOW : L_TT1P_scSF_PickAndPlaceHigh;
	XDONE : BOOL;
	XBUSY : BOOL;
	XACTIVE : BOOL;
	XAXESGROUPHOMED : BOOL;
	XINPOSITION : BOOL;
	XHWLIMITSWITCHACTIVE : BOOL;
	XSWLIMITSWITCHACTIVE : BOOL;
	AXHWLIMITSWITCHNEG : ARRAY [1..18] OF BOOL;
	AXHWLIMITSWITCHPOS : ARRAY [1..18] OF BOOL;
	AXSWLIMITSWITCHENABLE : ARRAY [1..18] OF BOOL;
	AXSWLIMITSWITCHACTIVE : ARRAY [1..18] OF BOOL;
	XPATHHOLD : BOOL;
	XGRIPPERCTRLACTIVE : BOOL;
	XPULSEGRIPPER : BOOL;
	LRSETPATHVELOUT : LREAL;
	LRPATHPREPARATIONTIME : LREAL;
	LRPRECALCPROFILETIME : LREAL;
	ALRACTAXISPOS : ARRAY [1..18] OF LREAL;
	ALRACTAXISVEL : ARRAY [1..18] OF LREAL;
	IPROFILEPOINTPASSED : INT;
	ISETPROFILENOOUT : INT;
	XPROFILEINPREPARATION : BOOL;
END_VAR
VAR_IN_OUT
	AXESGROUP : AXES_GROUP_KIN;
END_VAR
VAR
	TM_INT : _TM_PickAndPlaceHigh;
	PPAR : POINTER TO L_TT1P_scPar_PickAndPlaceHigh;
	PPAR_INT : POINTER TO L_TT1P_scPar_PickAndPlaceHigh;
	FB_LIMITDYNAMICSMAINAXES : L_MC4P_LimitDynamicsMainAxes;
	FB_LIMITDYNAMICSAUXAXES : L_MC4P_LimitDynamicsAuxAxes;
	AFB_HWLIMITAXIS : ARRAY [1..13] OF L_MC1P_HWLimitSwitchInterface;
END_VAR
END_FUNCTION_BLOCK

(* ---- L_TT1P_PICKANDPLACESTATE.fb ---- *)
FUNCTION_BLOCK L_TT1P_PICKANDPLACESTATE
VAR_INPUT
	XENABLEINTERNALCONTROL : BOOL;
	XENABLE : BOOL;
	SCCTRLAGBC : scCtrl_AGBC;
	XRESETERROR : BOOL;
	XREGULATORONALL : BOOL;
	XPATHSTOP : BOOL;
	XPATHHALT : BOOL;
	XSTOPALL : BOOL;
	SCPAR : L_TT1P_scPar_PickAndPlaceState;
	SCACCESSPOINTS : L_TT1P_scAP_PickAndPlaceState;
	XEXECUTEPICKANDPLACE : BOOL;
	XPATHINTERRUPT : BOOL;
	XGROUPHOMEEXECUTE : BOOL;
	AXHOMEABSSWITCH : ARRAY [1..12] OF BOOL;
	XGROUPENABLEHWLIMIT : BOOL;
	AXHWLIMITPOS : ARRAY [1..18] OF BOOL;
	AXHWLIMITNEG : ARRAY [1..18] OF BOOL;
	ESELECTAXIS : IDENT_IN_GROUP_REF;
	XJOGPOS : BOOL;
	XJOGNEG : BOOL;
	XABORT : BOOL;
	LROVERRIDE : LREAL := 1;
	XACKPATHHALT : BOOL;
END_VAR
VAR_OUTPUT
	XINTERNALCONTROLACTIVE : BOOL;
	ETMSTATE : L_TT1P_States := L_TT1P_States.INIT;
	SCSTATUSAGBC : scStatus_AGBC;
	XERROR : BOOL;
	XWARNING : BOOL;
	EERRORID : L_IE1P_Error;
	ASCERRORINFO : ARRAY [1..18] OF L_TT1P_scErrorInfo;
	XAXESENABLED : BOOL;
	XAXESGROUPENABLED : BOOL;
	SCSIGNALFLOW : L_TT1P_scSF_PickAndPlaceState;
	XDONE : BOOL;
	XBUSY : BOOL;
	XACTIVE : BOOL;
	XAXESGROUPHOMED : BOOL;
	XINPOSITION : BOOL;
	XHWLIMITSWITCHACTIVE : BOOL;
	XSWLIMITSWITCHACTIVE : BOOL;
	AXHWLIMITSWITCHNEG : ARRAY [1..18] OF BOOL;
	AXHWLIMITSWITCHPOS : ARRAY [1..18] OF BOOL;
	AXSWLIMITSWITCHENABLE : ARRAY [1..18] OF BOOL;
	AXSWLIMITSWITCHACTIVE : ARRAY [1..18] OF BOOL;
	XPATHHOLD : BOOL;
	XGRIPPERCTRLACTIVE : BOOL;
	XPULSEGRIPPER : BOOL;
	LRSETPATHVELOUT : LREAL;
	LRPATHPREPARATIONTIME : LREAL;
	LRPRECALCPROFILETIME : LREAL;
	ALRACTAXISPOS : ARRAY [1..18] OF LREAL;
	ALRACTAXISVEL : ARRAY [1..18] OF LREAL;
	IPROFILEPOINTPASSED : INT;
END_VAR
VAR_IN_OUT
	AXESGROUP : AXES_GROUP_KIN;
END_VAR
VAR
	TM_INT : _TM_PickAndPlaceStateExtension;
	PPAR : POINTER TO L_TT1P_scPar_PickAndPlaceState;
	PPAR_INT : POINTER TO L_TT1P_scPar_PickAndPlaceState;
	FB_LIMITDYNAMICSMAINAXES : L_MC4P_LimitDynamicsMainAxes;
	FB_LIMITDYNAMICSAUXAXES : L_MC4P_LimitDynamicsAuxAxes;
	AFB_HWLIMITAXIS : ARRAY [1..13] OF L_MC1P_HWLimitSwitchInterface;
END_VAR
END_FUNCTION_BLOCK

(* ---- L_TT1P_POSTRANSITION.fb ---- *)
FUNCTION_BLOCK L_TT1P_POSTRANSITION
VAR_INPUT
	LRPOSIN : LREAL;
	LRTRANSISTION : LREAL;
END_VAR
VAR_OUTPUT
	XERROR : BOOL;
	XTRANSITIONPOS : BOOL;
	XTRANSITIONNEG : BOOL;
	XTRANSITION : BOOL;
END_VAR
VAR_IN_OUT
	AXISDATA : AXIS_REF;
END_VAR
VAR
	LRDELTAPOSITION : LREAL;
	LRDELTAPOSITIONOLD : LREAL;
	L_MB1P_DIFFERENTIATE1 : L_MC2P_Differentiate;
	XINITDONE : BOOL;
END_VAR
END_FUNCTION_BLOCK

(* ---- L_TT1P_PROCESSCONTROL.fb ---- *)
FUNCTION_BLOCK L_TT1P_PROCESSCONTROL
VAR_INPUT
	XENABLE : BOOL;
	XSYNCFLYINGSAW : BOOL;
	XSYNCININSTANT : BOOL;
	XEXECUTEFIRSTCUT : BOOL;
	XRESUMETARGETPOS : BOOL;
	XRESET : BOOL;
	XTPNOTVALID : BOOL;
	XEXECUTEGAP : BOOL;
	XDONEPROFILE : BOOL;
	LRSLAVEPOSIN : LREAL;
	LRLOWERLIMIT : LREAL;
	LRUPPERLIMIT : LREAL;
	LRSTARTPOS : LREAL;
	LRPOSX1 : LREAL;
	LRVELX1 : LREAL;
	LRACCX1 : LREAL;
	LRTASKCYCLE : LREAL;
END_VAR
VAR_OUTPUT
	XEXECUTEPROFILE : BOOL;
	XAUXEXECUTEPROFILE : BOOL;
	XSYNCPOSOUT : BOOL;
	LRPOSX2 : LREAL;
	LRVELX2 : LREAL;
	LRACCX2 : LREAL;
	XCUTTINGACTIVE : BOOL;
	LRTOLERANCE : LREAL;
END_VAR
VAR
	XEXECUTEPROFILE_INT : BOOL;
	XSYNC_INT : BOOL;
	WSTEPPER : WORD;
	XEXECUTEGAP_OLD : BOOL;
	XRESET_OLD : BOOL;
	XSYNCININSTANT_OLD : BOOL;
	XENABLE_OLD : BOOL;
	LRSTARTTHRESHOLD : LREAL;
	XRESUMETARGETPOS_OLD : BOOL;
	XEXECUTEFIRSTCUT_OLD : BOOL;
END_VAR
END_FUNCTION_BLOCK

(* ---- L_TT1P_REGISTERCONTROLBASE.fb ---- *)
FUNCTION_BLOCK L_TT1P_REGISTERCONTROLBASE
VAR_INPUT
	XENABLEINTERNALCONTROL : BOOL;
	XENABLE : BOOL;
	SCCTRLABC : scCtrl_ABC;
	XRESETERROR : BOOL;
	XREGULATORON : BOOL;
	XSTOP : BOOL;
	XHALT : BOOL;
	SCPAR : L_TT1P_scPar_RegisterControlBase;
	SCACCESSPOINTS : L_TT1P_scAP_RegisterControlBase;
	XJOGPOS : BOOL;
	XJOGNEG : BOOL;
	XHOMEEXECUTE : BOOL;
	XHOMEABSSWITCH : BOOL;
	LRSETOFFSETMASTER : LREAL;
	LRSETOFFSETSLAVE : LREAL;
	XTRIMPOS : BOOL;
	XTRIMNEG : BOOL;
	XSYNCPOS : BOOL;
	XSYNCINSTANT : BOOL;
	XSYNCOUTINSTANT : BOOL;
	XSYNCPOSRESTORE : BOOL;
	XMARKRECEIVE : BOOL;
	LRACTMARKPOSIN : LREAL;
	LRCYCPOSEXTENCODER : LREAL;
	XLOADREGPOS : BOOL;
	LRLOADREGPOS : LREAL;
END_VAR
VAR_OUTPUT
	XINTERNALCONTROLACTIVE : BOOL;
	ETMSTATE : L_TT1P_States := L_TT1P_States.INIT;
	SCSTATUSABC : scStatus_ABC;
	XERROR : BOOL;
	XWARNING : BOOL;
	EERRORID : L_IE1P_Error;
	SCERRORINFO : L_TT1P_scErrorInfo;
	XAXISENABLED : BOOL;
	SCSIGNALFLOW : L_TT1P_scSF_RegisterControlBase;
	XDONE : BOOL;
	XBUSY : BOOL;
	XISHOMED : BOOL;
	LRACTVEL : LREAL;
	LRACTPOS : LREAL;
	LROFFSET : LREAL;
	LROFFSETTRIM : LREAL;
	LROFFSETTOTAL : LREAL;
	XSYNCHRONISED : BOOL;
	XACCDECSYNC : BOOL;
	LROFFSETSYNCPOS : LREAL;
	LRSETREGPOSOUT : LREAL;
	LRMARKSENSORPOS : LREAL;
	LRACTMARKERROR : LREAL;
	LRACTMARKDIST : LREAL;
	XMARKRECEIVED : BOOL;
	LRREGMARKPOS : LREAL;
	XCORRACTIVE : BOOL;
	XCORRLIMITED : BOOL;
END_VAR
VAR_IN_OUT
	MASTERAXIS : AXIS_REF;
	SLAVEAXIS : AXIS_REF;
END_VAR
VAR
	TM_INT : _TM_RegisterControlBase;
	PPARREG : POINTER TO L_TT1P_scPar_RegisterControlBase;
	PPARREG_INT : POINTER TO L_TT1P_scPar_RegisterControlBase;
	SCSIGNALFLOWES : _scSF_TM_ElectricalShaftPosHigh;
	LROFFSETMASTER : LREAL := 0;
END_VAR
END_FUNCTION_BLOCK

(* ---- L_TT1P_REGISTERCONTROLSTATE.fb ---- *)
FUNCTION_BLOCK L_TT1P_REGISTERCONTROLSTATE
VAR_INPUT
	XENABLEINTERNALCONTROL : BOOL;
	XENABLE : BOOL;
	SCCTRLABC : scCtrl_ABC;
	XRESETERROR : BOOL;
	XREGULATORON : BOOL;
	XSTOP : BOOL;
	XHALT : BOOL;
	SCPAR : L_TT1P_scPar_RegisterControlState;
	SCACCESSPOINTS : L_TT1P_scAP_RegisterControlState;
	XJOGPOS : BOOL;
	XJOGNEG : BOOL;
	XHOMEEXECUTE : BOOL;
	XHOMEABSSWITCH : BOOL;
	LRSETOFFSETMASTER : LREAL;
	LRSETOFFSETSLAVE : LREAL;
	XTRIMPOS : BOOL;
	XTRIMNEG : BOOL;
	XSYNCPOS : BOOL;
	XSYNCINSTANT : BOOL;
	XSYNCOUTINSTANT : BOOL;
	XSYNCPOSRESTORE : BOOL;
	XMARKRECEIVE : BOOL;
	LRACTMARKPOSIN : LREAL;
	LRCYCPOSEXTENCODER : LREAL;
	XLOADREGPOS : BOOL;
	LRLOADREGPOS : LREAL;
	XGEARFACTORCORR : BOOL;
	XGEARFACTORCORRHOLD : BOOL;
	XTEACHMARKWINDOW : BOOL;
END_VAR
VAR_OUTPUT
	XINTERNALCONTROLACTIVE : BOOL;
	ETMSTATE : L_TT1P_States := L_TT1P_States.INIT;
	SCSTATUSABC : scStatus_ABC;
	XERROR : BOOL;
	XWARNING : BOOL;
	EERRORID : L_IE1P_Error;
	SCERRORINFO : L_TT1P_scErrorInfo;
	XAXISENABLED : BOOL;
	SCSIGNALFLOW : L_TT1P_scSF_RegisterControlState;
	XDONE : BOOL;
	XBUSY : BOOL;
	XISHOMED : BOOL;
	LRACTVEL : LREAL;
	LRACTPOS : LREAL;
	LROFFSET : LREAL;
	LROFFSETTRIM : LREAL;
	LROFFSETTOTAL : LREAL;
	XSYNCHRONISED : BOOL;
	XACCDECSYNC : BOOL;
	LROFFSETSYNCPOS : LREAL;
	LRSETREGPOSOUT : LREAL;
	LRMARKSENSORPOS : LREAL;
	LRACTMARKERROR : LREAL;
	LRACTMARKDIST : LREAL;
	XMARKRECEIVED : BOOL;
	LRREGMARKPOS : LREAL;
	XCORRACTIVE : BOOL;
	XCORRLIMITED : BOOL;
	XMARKWINDOWOPEN : BOOL;
	XMARKOUTOFWINDOW : BOOL;
	XMARKNOTDETECTED : BOOL;
	XMARKWINDOWTEACHED : BOOL;
	LRAVERAGEGEARFACTORCORR : LREAL;
	XGEARFACTORCORRLIMITED : BOOL;
END_VAR
VAR_IN_OUT
	MASTERAXIS : AXIS_REF;
	SLAVEAXIS : AXIS_REF;
END_VAR
VAR
	TM_INT : _TM_RegisterControlState;
	PPARREG : POINTER TO L_TT1P_scPar_RegisterControlState;
	PPARREG_INT : POINTER TO L_TT1P_scPar_RegisterControlState;
	SCSIGNALFLOWES : _scSF_TM_ElectricalShaftPosHigh;
	LROFFSETMASTER : LREAL := 0;
END_VAR
END_FUNCTION_BLOCK

METHOD GET_LRMARKSTACKLENGTH : LREAL
END_METHOD

(* ---- L_TT1P_SMARTTRACKBASE.fb ---- *)
FUNCTION_BLOCK L_TT1P_SMARTTRACKBASE
VAR_INPUT
	XENABLEINTERNALCONTROL : BOOL;
	XENABLE : BOOL;
	SCCTRLABC : scCtrl_ABC;
	XRESETERROR : BOOL;
	XREGULATORON : BOOL;
	XSTOP : BOOL;
	XHALT : BOOL;
	SCPAR : L_TT1P_scPar_SmartTrackBase;
	SCACCESSPOINTS : L_TT1P_scAP_SmartTrackBase;
	XJOGPOS : BOOL;
	XJOGNEG : BOOL;
	XSYNCVEL : BOOL;
	XPRODUCTEDGERISE : BOOL;
	XPRODUCTEDGEFALL : BOOL;
	LRACTPRODUCTEDGEPOSIN : LREAL;
END_VAR
VAR_OUTPUT
	XINTERNALCONTROLACTIVE : BOOL;
	ETMSTATE : L_TT1P_States := L_TT1P_States.INIT;
	SCSTATUSABC : scStatus_ABC;
	XERROR : BOOL;
	XWARNING : BOOL;
	EERRORID : L_IE1P_Error;
	SCERRORINFO : L_TT1P_scErrorInfo;
	XAXISENABLED : BOOL;
	SCSIGNALFLOW : L_TT1P_scSF_SmartTrackBase;
	XDONE : BOOL;
	XBUSY : BOOL;
	LRACTPOS : LREAL;
	LRACTVEL : LREAL;
	LRACTFOLLOWINGERROR : LREAL;
	XPRODUCTRECEIVED : BOOL;
	LRACTPRODUCTERROR : LREAL;
	LRACTPRODUCTERRORLIMITED : LREAL;
	LRMASTERPOSEDGERISE : LREAL;
	XCORRACTIVE : BOOL;
	XCORRLIMITED : BOOL;
END_VAR
VAR_IN_OUT
	MASTERAXIS : AXIS_REF;
	SLAVEAXIS : AXIS_REF;
END_VAR
VAR
	TM_INT : _TM_SmartTrackBase;
	PPAR : POINTER TO L_TT1P_scPar_SmartTrackBase;
	PPAR_INT : POINTER TO L_TT1P_scPar_SmartTrackBase;
	XHOMEEXECUTE : BOOL;
	XHOMEABSSWITCH : BOOL;
	XISHOMED : BOOL;
END_VAR
END_FUNCTION_BLOCK

(* ---- L_TT1P_SMARTTRACKSTATE.fb ---- *)
FUNCTION_BLOCK L_TT1P_SMARTTRACKSTATE
VAR_INPUT
	XENABLEINTERNALCONTROL : BOOL;
	XENABLE : BOOL;
	SCCTRLABC : scCtrl_ABC;
	XRESETERROR : BOOL;
	XREGULATORON : BOOL;
	XSTOP : BOOL;
	XHALT : BOOL;
	SCPAR : L_TT1P_scPar_SmartTrackState;
	SCACCESSPOINTS : L_TT1P_scAP_SmartTrackState;
	XJOGPOS : BOOL;
	XJOGNEG : BOOL;
	XSYNCVEL : BOOL;
	XPRODUCTEDGERISE : BOOL;
	XPRODUCTEDGEFALL : BOOL;
	LRACTPRODUCTEDGEPOSIN : LREAL;
	DATABUSIN : ITF_DataBus;
END_VAR
VAR_OUTPUT
	XINTERNALCONTROLACTIVE : BOOL;
	ETMSTATE : L_TT1P_States := L_TT1P_States.INIT;
	SCSTATUSABC : scStatus_ABC;
	XERROR : BOOL;
	XWARNING : BOOL;
	EERRORID : L_IE1P_Error;
	SCERRORINFO : L_TT1P_scErrorInfo;
	XAXISENABLED : BOOL;
	SCSIGNALFLOW : L_TT1P_scSF_SmartTrackState;
	XDONE : BOOL;
	XBUSY : BOOL;
	LRACTPOS : LREAL;
	LRACTVEL : LREAL;
	LRACTFOLLOWINGERROR : LREAL;
	XPRODUCTRECEIVED : BOOL;
	LRACTPRODUCTERROR : LREAL;
	LRACTPRODUCTERRORLIMITED : LREAL;
	LRMASTERPOSEDGERISE : LREAL;
	XCORRACTIVE : BOOL;
	XCORRLIMITED : BOOL;
	DATABUSOUT : ITF_DataBus;
	XCOMMUNICATIONVALID : BOOL;
	XMASTER : BOOL;
	XSLAVE : BOOL;
	BYSMARTTRACKNO : BYTE;
	LRDISTTOOUTFEED : LREAL;
END_VAR
VAR_IN_OUT
	MASTERAXIS : AXIS_REF;
	SLAVEAXIS : AXIS_REF;
END_VAR
VAR
	TM_INT : _TM_SmartTrackState;
	PPAR : POINTER TO L_TT1P_scPar_SmartTrackState;
	PPAR_INT : POINTER TO L_TT1P_scPar_SmartTrackState;
	XHOMEEXECUTE : BOOL;
	XHOMEABSSWITCH : BOOL;
	XISHOMED : BOOL;
END_VAR
END_FUNCTION_BLOCK

(* ---- L_TT1P_STACKERCRANEAXISCONTROLBASE.fb ---- *)
FUNCTION_BLOCK L_TT1P_STACKERCRANEAXISCONTROLBASE
VAR_INPUT
	XENABLEINTERNALCONTROL : BOOL;
	XENABLE : BOOL;
	SCCTRLABC : scCtrl_ABC;
	XRESETERROR : BOOL;
	XREGULATORON : BOOL;
	XSTOP : BOOL;
	XHALT : BOOL;
	SCPAR : L_TT1P_scPar_StackerCraneAxisControlBase;
	DATABUSIN : ITF_DataBus;
	EADDRESS : L_TT1P_StackerCraneAddress := 0;
	SCACCESSPOINTS : L_TT1P_scAP_StackerCraneAxisControlBase;
	XJOGPOS : BOOL;
	XJOGNEG : BOOL;
	XHOMEEXECUTE : BOOL;
	XHOMEABSSWITCH : BOOL;
	LROVERRIDE : LREAL := 1.0;
	XOSCCOMP : BOOL;
	LROSCCOMPPOSSCALED : LREAL;
	LROSCCOMPLOADSCALED : LREAL;
	XEXECUTEBRAKETEST : BOOL;
	XEXECUTEBRAKEGRINDIN : BOOL;
END_VAR
VAR_OUTPUT
	XINTERNALCONTROLACTIVE : BOOL;
	ETMSTATE : L_TT1P_States;
	SCSTATUSABC : scStatus_ABC;
	XERROR : BOOL;
	XWARNING : BOOL;
	EERRORID : L_IE1P_Error;
	SCERRORINFO : L_TT1P_scErrorInfo;
	XAXISENABLED : BOOL;
	SCSIGNALFLOW : L_TT1P_scSF_StackerCraneAxisControlBase;
	XAXISREADY : BOOL;
	XISHOMED : BOOL;
	XDONE : BOOL;
	XBUSY : BOOL;
	XCOMMANDABORTED : BOOL;
	XINPOSITION : BOOL;
	ECONTROLMODE : L_MC1P_ControlMode;
	LRACTVEL : LREAL;
	LRACTPOS : LREAL;
	XOSCCOMPACTIVE : BOOL;
END_VAR
VAR_IN_OUT
	AXIS : AXIS_REF;
END_VAR
VAR
	TM_INT : _TM_StackerCraneAxisControlBase;
END_VAR
END_FUNCTION_BLOCK

(* ---- L_TT1P_STACKERCRANEHEADCONTROLBASE.fb ---- *)
FUNCTION_BLOCK L_TT1P_STACKERCRANEHEADCONTROLBASE
VAR_INPUT
	XENABLEINTERNALCONTROL : BOOL;
	XENABLE : BOOL;
	XRESETERROR : BOOL;
	XSTOPALL : BOOL;
	SCPAR : L_TT1P_scPar_StackerCraneHeadControlBase;
	XEXECUTEPROFILEX : BOOL;
	XEXECUTEPROFILEY : BOOL;
	XMAINTENANCEMODE : BOOL;
END_VAR
VAR_OUTPUT
	DATABUSOUT : ITF_DataBus;
	XINTERNALCONTROLACTIVE : BOOL;
	ETMSTATE : L_TT1P_States;
	XERROR : BOOL;
	XWARNING : BOOL;
	EERRORID : L_IE1P_Error;
	ASCERRORINFO : ARRAY [1..6] OF L_TT1P_scErrorInfo;
	XAXESENABLED : BOOL;
	SCSIGNALFLOW : L_TT1P_scSF_StackerCraneHeadControlBase;
	XAXESREADY : BOOL;
	XAXESHOMED : BOOL;
	XPROFILEXDONE : BOOL;
	XPROFILEYDONE : BOOL;
	XPROFILEXBUSY : BOOL;
	XPROFILEYBUSY : BOOL;
END_VAR
VAR
	TM_INT : _TM_StackerCraneHeadControlBase;
END_VAR
END_FUNCTION_BLOCK

(* ---- L_TT1P_TABLEPOSITIONINGBASE.fb ---- *)
FUNCTION_BLOCK L_TT1P_TABLEPOSITIONINGBASE
VAR_INPUT
	XENABLEINTERNALCONTROL : BOOL;
	XENABLE : BOOL;
	SCCTRLABC : scCtrl_ABC;
	XRESETERROR : BOOL;
	XREGULATORON : BOOL;
	XSTOP : BOOL;
	XHALT : BOOL;
	SCPAR : L_TT1P_scPar_TablePositioningBase;
	SCACCESSPOINTS : L_TT1P_scAP_TablePositioningBase;
	XJOGPOS : BOOL;
	XJOGNEG : BOOL;
	XHOMEEXECUTE : BOOL;
	XHOMEABSSWITCH : BOOL;
	XRESETHOMEPOSITION : BOOL;
	XHWLIMITPOS : BOOL;
	XHWLIMITNEG : BOOL;
	EPROFILENUMBER : L_TT1P_ProfileNumber;
	XEXECUTEPOSITIONING : BOOL;
	XABORTPOSITIONING : BOOL;
	XFINISHPOSITIONING : BOOL;
	XTPRECEIVE : BOOL;
	LRACTTPPOSITION : LREAL;
	LRCYCPOSEXTENCODER : LREAL;
	LRSETTORQUELIMITPOS : LREAL;
	LRSETTORQUELIMITNEG : LREAL;
	LRSETOVERRIDEVEL : LREAL;
	LRSETOVERRIDEACCDEC : LREAL;
	LRSETOVERRIDEJERK : LREAL;
END_VAR
VAR_OUTPUT
	XINTERNALCONTROLACTIVE : BOOL;
	ETMSTATE : L_TT1P_States := L_TT1P_States.INIT;
	SCSTATUSABC : scStatus_ABC;
	XERROR : BOOL;
	XWARNING : BOOL;
	EERRORID : L_IE1P_Error;
	SCERRORINFO : L_TT1P_scErrorInfo;
	XAXISENABLED : BOOL;
	SCSIGNALFLOW : L_TT1P_scSF_TablePositioningBase;
	XDONE : BOOL;
	XBUSY : BOOL;
	XISHOMED : BOOL;
	LRACTPOS : LREAL;
	LRACTVEL : LREAL;
	LRACTFOLLOWINGERROR : LREAL;
	XPOSITIONINGACTIVE : BOOL;
	XPOSITIONINGDONE : BOOL;
	XDRIVEINTARGET : BOOL;
	XTPRECEIVED : BOOL;
	XTPMISSED : BOOL;
	XTPOUTOFWINDOW : BOOL;
	EACTIVEPROFILE : L_TT1P_ProfileNumber;
END_VAR
VAR_IN_OUT
	AXIS : AXIS_REF;
END_VAR
VAR
	TM_INT : _TM_TablePositioningBase;
	PPAR : POINTER TO L_TT1P_scPar_TablePositioningBase;
	PPAR_INT : POINTER TO L_TT1P_scPar_TablePositioningBase;
END_VAR
END_FUNCTION_BLOCK

(* ---- L_TT1P_VIRTUALMASTERBASE.fb ---- *)
FUNCTION_BLOCK L_TT1P_VIRTUALMASTERBASE
VAR_INPUT
	XENABLEINTERNALCONTROL : BOOL;
	XENABLE : BOOL;
	SCCTRLABC : scCtrl_ABC;
	XRESETERROR : BOOL;
	XREGULATORON : BOOL;
	XSTOP : BOOL;
	XHALT : BOOL;
	SCPAR : L_TT1P_scPar_VirtualMasterBase;
	XCONTINUOUS : BOOL;
	XCYCLE : BOOL;
	XLOADSTARTPOS : BOOL;
	XJOGPOS : BOOL;
	XJOGNEG : BOOL;
	LRSETVEL : LREAL := 10;
	LRSTARTPOS : LREAL;
	LRTARGETPOS : LREAL;
END_VAR
VAR_OUTPUT
	XINTERNALCONTROLACTIVE : BOOL;
	ETMSTATE : L_TT1P_States := L_TT1P_States.INIT;
	SCSTATUSABC : scStatus_ABC;
	XERROR : BOOL;
	XWARNING : BOOL;
	EERRORID : L_IE1P_Error;
	SCERRORINFO : L_TT1P_scErrorInfo;
	XAXISENABLED : BOOL;
	XBUSY : BOOL;
	XINTARGET : BOOL;
	LRACTPOS : LREAL;
	LRACTVEL : LREAL;
	LRSETPOSOUT : LREAL;
	LRSETVELOUT : LREAL;
END_VAR
VAR_IN_OUT
	VIRTUALAXIS : AXIS_REF;
END_VAR
VAR
	TM_INT : _TM_VirtualMasterBase;
	PPAR : POINTER TO L_TT1P_scPar_VirtualMasterBase;
	PPAR_INT : POINTER TO L_TT1P_scPar_VirtualMasterBase;
	XDONE : BOOL;
	XHOMEEXECUTE : BOOL;
	XHOMEABSSWITCH : BOOL;
	XISHOMED : BOOL;
	SCACCESSPOINTS : _scAP_TM_MotionControl;
	SCSIGNALFLOW : _scSF_TM_MotionControl;
END_VAR
END_FUNCTION_BLOCK

(* ---- L_TT1P_VIRTUALMASTERHIGH.fb ---- *)
FUNCTION_BLOCK L_TT1P_VIRTUALMASTERHIGH
VAR_INPUT
	XENABLEINTERNALCONTROL : BOOL;
	XENABLE : BOOL;
	SCCTRLABC : scCtrl_ABC;
	XRESETERROR : BOOL;
	XREGULATORON : BOOL;
	XSTOP : BOOL;
	XHALT : BOOL;
	SCPAR : L_TT1P_scPar_VirtualMasterHigh;
	MASTERAXIS : L_MC1P_IAXIS_REF_MASTERVALUES;
	XCONTINUOUS : BOOL;
	XCYCLE : BOOL;
	XLOADSTARTPOS : BOOL;
	XJOGPOS : BOOL;
	XJOGNEG : BOOL;
	LRSETVEL : LREAL := 10;
	LRSTARTPOS : LREAL;
	LRTARGETPOS : LREAL;
	XSYNCMASTERAXIS : BOOL;
END_VAR
VAR_OUTPUT
	XINTERNALCONTROLACTIVE : BOOL;
	ETMSTATE : L_TT1P_States := L_TT1P_States.INIT;
	SCSTATUSABC : scStatus_ABC;
	XERROR : BOOL;
	XWARNING : BOOL;
	EERRORID : L_IE1P_Error;
	SCERRORINFO : L_TT1P_scErrorInfo;
	XAXISENABLED : BOOL;
	XBUSY : BOOL;
	XINTARGET : BOOL;
	LRACTPOS : LREAL;
	LRACTVEL : LREAL;
	LRSETPOSOUT : LREAL;
	LRSETVELOUT : LREAL;
	XACCDECSYNC : BOOL;
	XSYNCHRONISED : BOOL;
END_VAR
VAR_IN_OUT
	VIRTUALAXIS : AXIS_REF;
END_VAR
VAR
	TM_INT : _TM_VirtualMasterHigh;
	PPAR : POINTER TO L_TT1P_scPar_VirtualMasterHigh;
	PPAR_INT : POINTER TO L_TT1P_scPar_VirtualMasterHigh;
	XDONE : BOOL;
	XHOMEEXECUTE : BOOL;
	XHOMEABSSWITCH : BOOL;
	XISHOMED : BOOL;
	SCACCESSPOINTS : _scAP_TM_MotionControl;
	SCSIGNALFLOW : _scSF_TM_MotionControl;
END_VAR
END_FUNCTION_BLOCK

(* ---- L_TT1P_VIRTUALMASTERSTATE.fb ---- *)
FUNCTION_BLOCK L_TT1P_VIRTUALMASTERSTATE
VAR_INPUT
	XENABLEINTERNALCONTROL : BOOL;
	XENABLE : BOOL;
	SCCTRLABC : scCtrl_ABC;
	XRESETERROR : BOOL;
	XREGULATORON : BOOL;
	XSTOP : BOOL;
	XHALT : BOOL;
	SCPAR : L_TT1P_scPar_VirtualMasterState;
	MASTERAXIS : L_MC1P_IAXIS_REF_MASTERVALUES;
	XCONTINUOUS : BOOL;
	XCYCLE : BOOL;
	XLOADSTARTPOS : BOOL;
	XJOGPOS : BOOL;
	XJOGNEG : BOOL;
	LRSETVEL : LREAL := 10;
	LRSTARTPOS : LREAL;
	LRTARGETPOS : LREAL;
	XSYNCMASTERAXIS : BOOL;
END_VAR
VAR_OUTPUT
	XINTERNALCONTROLACTIVE : BOOL;
	ETMSTATE : L_TT1P_States := L_TT1P_States.INIT;
	SCSTATUSABC : scStatus_ABC;
	XERROR : BOOL;
	XWARNING : BOOL;
	EERRORID : L_IE1P_Error;
	SCERRORINFO : L_TT1P_scErrorInfo;
	XAXISENABLED : BOOL;
	XBUSY : BOOL;
	XINTARGET : BOOL;
	LRACTPOS : LREAL;
	LRACTVEL : LREAL;
	LRSETPOSOUT : LREAL;
	LRSETVELOUT : LREAL;
	XACCDECSYNC : BOOL;
	XSYNCHRONISED : BOOL;
END_VAR
VAR_IN_OUT
	VIRTUALAXIS : AXIS_REF;
END_VAR
VAR
	TM_INT : _TM_VirtualMasterState;
	PPAR : POINTER TO L_TT1P_scPar_VirtualMasterState;
	PPAR_INT : POINTER TO L_TT1P_scPar_VirtualMasterState;
	XDONE : BOOL;
	XHOMEEXECUTE : BOOL;
	XHOMEABSSWITCH : BOOL;
	XISHOMED : BOOL;
	SCACCESSPOINTS : _scAP_TM_MotionControl;
	SCSIGNALFLOW : _scSF_TM_MotionControl;
END_VAR
END_FUNCTION_BLOCK
